(* IEC 61131-3 sources: daoli-st-library/DL_Device (part 23) *)

(* ---- FB_DL_GreaseLubeTimer.st ---- *)
(*
  Name        : FB_DL_GreaseLubeTimer
  Category    : DL_Device
  Version     : 1.0.0
  Purpose     : 加脂保养窗：运行小时数与动作循环数双触发（任一达限即报「该加脂」，先到先报），保养完成后复位清零重计；/ Grease lubrication window: running hours and cycle count both trigger (whichever reaches its limit first reports), cleared and restarted after maintenance
  溯源        : 借 t2-8 ◐/自研 的分类/参数域组织，clean-room 实现
  Boundary    : ① 组态闸：小时限/循环限任一 < 0 → 锁存故障（两限可独立为 0 表示该源不触发，但不可为负）；
                ② 运行小时用 1 s 自复位 TON 节拍累计（IN 串 eRun 相位 + bRunning，R188/族③），段 0 无 IF 包裹；
                ③ 双触发独立判据独立归因（R190）：eHoursFirst / eCyclesFirst 各自成因，同拍同到按小时优先归因（不共用成员）；
                ④ 秒计数饱和累加（R28 防回绕），循环数沿计数净额 +1 饱和；
                ⑤ bLubeDue 锁存至复位沿或 bLubeDone 沿（保养完成脉冲，唯一业务清零路径）；
                ⑥ 本件只报保养到期，不执行加脂动作（属主边界）。
*)
TYPE E_DL_GltState :
(
    eIdle  := 0,                             (* 未使能 / Disabled *)
    eRun   := 10,                            (* 保养窗计时计数运行 / Accumulating *)
    eFault := 90                             (* 故障锁存相 / Fault latched *)
);
END_TYPE

TYPE E_DL_GltCause :
(
    eNone        := 0,                       (* 无故障成因 / No cause *)
    eCfgIllegal  := 1,                       (* 组态非法：时限/循环限越域 / Illegal config *)
    eHoursFirst  := 2,                       (* 运行小时先达限（先到先报） / Hours limit reached first *)
    eCyclesFirst := 3,                       (* 动作循环先达限（先到先报） / Cycles limit reached first *)
    ePhaseBad    := 4                        (* 非法相位兜底 / Illegal phase fallback *)
);
END_TYPE

FUNCTION_BLOCK FB_DL_GreaseLubeTimer
VAR_INPUT
    bRunning   : BOOL := FALSE;              (* 设备运行电平（运行小时累计门控）[-] / Equipment running level *)
    bCyclePulse: BOOL := FALSE;              (* 动作循环脉冲（上升沿计一次）[-] / One action-cycle pulse *)
    fHoursLimit: REAL := 2000.0;             (* 运行小时触发限，域 >= 0（0 = 该源禁用）[h] / Hours trigger limit, >= 0 *)
    nCycleLimit: UDINT := 100000;            (* 循环数触发限，域 >= 0（0 = 该源禁用）[次] / Cycle trigger limit, >= 0 *)
    bLubeDone  : BOOL := FALSE;              (* 保养完成脉冲（业务清零路径，重开保养窗）[-] / Maintenance done pulse *)
    bEnable    : BOOL := TRUE;               (* 使能 [-] / Enable *)
    bReset     : BOOL := FALSE;              (* 复位命令，上升沿清累计与故障 [-] / Reset command *)
END_VAR
VAR_OUTPUT
    fRunHours  : REAL;                       (* 累计运行小时（窗内）[h] / Accumulated running hours *)
    nCycles    : UDINT;                      (* 累计动作循环数（窗内，饱和）[次] / Accumulated cycles, saturated *)
    bLubeDue   : BOOL;                       (* 加脂到期锁存（复位沿或保养完成沿清）[-] / Lubrication due latched *)
    eState     : E_DL_GltState;              (* 状态出口 / State outlet *)
    eCause     : E_DL_GltCause;              (* 成因出口（R190 双触发独立归因） / Cause outlet *)
    bError     : BOOL;                       (* 故障锁存标志 [-] / Fault latch flag *)
END_VAR
VAR
    _eState  : E_DL_GltState := E_DL_GltState.eIdle;     (* 内部相位（CASE 唯一写入目标） / Internal phase *)
    _eCause  : E_DL_GltCause := E_DL_GltCause.eNone;     (* 故障成因锁存量 / Latched cause *)
    rtCycle  : R_TRIG;                       (* 循环脉冲沿实例，段 0 无条件调用 / Cycle pulse edge *)
    rtLube   : R_TRIG;                       (* 保养完成沿实例，段 0 无条件调用 / Lube-done edge instance *)
    rtReset  : R_TRIG;                       (* 复位沿实例，段 0 无条件调用 / Reset edge instance *)
    tonTick  : TON;                          (* 1 s 节拍计时器（自复位，IN 串相位 + 运行电平） / 1 s tick timer *)
    _bFault  : BOOL;                         (* 故障锁存位 / Latched fault bit *)
    _bCfgBad : BOOL;                         (* 组态非法当拍量 / Illegal config this scan *)
    _fSec    : REAL;                         (* 窗内累计运行秒数（节拍累加）[s] / Accumulated seconds *)
    _fHoursI : REAL;                         (* 运行小时中间量（秒→小时换算）[h] / Hours intermediate *)
    _bDueI   : BOOL;                         (* 到期内部量（锁存副本源）[-] / Due internal, source of latch *)
END_VAR
VAR CONSTANT
    DL_GLT_EPS    : REAL  := 1.0E-6;         (* 判零容差 [-] / Epsilon *)
    DL_GLT_CNTMAX : UDINT := 4294967295;     (* 循环计数饱和上限（R28）[-] / Cycle count saturation cap *)
    DL_GLT_SECMAX : REAL  := 3.0E9;          (* 秒累计上限（防 REAL 有效位耗尽，约 95 年）[s] / Seconds accumulation cap *)
    DL_GLT_H2S    : REAL  := 3600.0;         (* 小时→秒换算常量（乘性常量）[-] / Hours to seconds factor *)
END_VAR

(* —— 段 0：当拍判据派生 + 实例无条件刷新（R228A；R_TRIG/TON 全在段 0，无 IF 包裹） —— *)
_bCfgBad := (fHoursLimit < 0.0) OR (nCycleLimit < 0);                          (* 两触发限非负闸（0 = 禁用该源，合法） / Limits non-negative gates *)
rtCycle(CLK := bCyclePulse);                                                   (* 循环沿每拍必调 / Cycle edge every scan *)
rtLube(CLK := bLubeDone);                                                      (* 保养完成沿每拍必调 / Done edge every scan *)
rtReset(CLK := bReset);                                                        (* 复位沿每拍必调 / Reset edge every scan *)
tonTick(IN := (_eState = E_DL_GltState.eRun) AND bRunning AND NOT tonTick.Q, PT := T#1S);   (* 1 s 节拍自复位（R188）+ eRun 相位与运行电平闸 / 1 s tick with phase and run gates *)

(* —— 段 1：单拍量预清零（R107） —— *)
_bDueI := FALSE;                                                               (* 到期内部量预清（判据拍重算） / Due internal preset *)
_fHoursI := 0.0;                                                               (* 小时中间量预清 / Hours intermediate preset *)

(* —— 段 2：复位沿处理（作用域：清故障 + 清累计 + 清到期 + 迁 eIdle，R283 逐项声明） —— *)
IF rtReset.Q THEN
    _bFault := FALSE;                                                          (* 清故障锁存 / Clear fault *)
    _eCause := E_DL_GltCause.eNone;                                            (* 清成因 / Clear cause *)
    _fSec := 0.0;                                                              (* 清秒累计 / Clear seconds *)
    nCycles := 0;                                                              (* 清循环计数出口 / Clear cycles outlet *)
    bLubeDue := FALSE;                                                         (* 清到期锁存出口 / Clear due outlet *)
    _eState := E_DL_GltState.eIdle;                                            (* 迁未使能相 / Back to idle *)
END_IF

(* —— 段 3：组态故障锁存（锁存至复位沿，R189） —— *)
IF _bCfgBad AND NOT _bFault THEN
    _bFault := TRUE;                                                           (* 锁存故障位 / Latch fault *)
    _eCause := E_DL_GltCause.eCfgIllegal;                                      (* 成因：组态非法 / Cause: illegal config *)
    _eState := E_DL_GltState.eFault;                                           (* 同步迁故障相 / Migrate to fault *)
END_IF

(* —— 段 4：CASE 主状态机（ELSE 兜底迁 eFault，红线 6） —— *)
CASE _eState OF
    E_DL_GltState.eIdle:                                                       (* 未使能：不累计，出口确定值 / Disabled *)
        _fSec := 0.0;                                                          (* 失能清秒累计（防隐性回夹） / Clear seconds *)
        fRunHours := 0.0;                                                      (* 失能清小时出口 / Clear hours outlet *)
        nCycles := 0;                                                          (* 失能清循环出口 / Clear cycles outlet *)
        bLubeDue := FALSE;                                                     (* 失能清到期出口 / Clear due outlet *)
        IF bEnable AND NOT _bFault THEN
            _eState := E_DL_GltState.eRun;                                     (* 使能进入累计 / Enter accumulating *)
        END_IF
    E_DL_GltState.eRun:                                                        (* 累计相：小时 + 循环双源 / Accumulating *)
        IF NOT bEnable THEN
            _eState := E_DL_GltState.eIdle;                                    (* 失能回未使能 / Back to idle *)
        ELSE
            IF rtLube.Q THEN                                                   (* 保养完成沿：业务清零重开窗（唯一业务清零路径） / Done edge: clear and reopen window *)
                _fSec := 0.0;                                                  (* 清秒累计 / Clear seconds *)
                nCycles := 0;                                                  (* 清循环计数 / Clear cycles *)
                bLubeDue := FALSE;                                             (* 清到期锁存 / Clear due latch *)
                _eCause := E_DL_GltCause.eNone;                                (* 成因复位 / Cause reset *)
            END_IF
            IF tonTick.Q THEN                                                  (* 1 s 节拍到点：秒累计 +1 / Tick elapsed: +1 second *)
                IF _fSec < DL_GLT_SECMAX THEN
                    _fSec := _fSec + 1.0;                                      (* 秒累计（饱和防有效位耗尽，R28） / Seconds accumulate, capped *)
                END_IF
            END_IF
            IF rtCycle.Q THEN                                                  (* 动作循环沿：循环计数 +1 / Cycle edge: +1 *)
                IF nCycles < DL_GLT_CNTMAX THEN
                    nCycles := nCycles + 1;                                    (* 循环计数净额 +1（饱和防回绕） / Net +1, saturated *)
                END_IF
            END_IF
            _fHoursI := _fSec / DL_GLT_H2S;                                    (* 秒→小时换算（除子为常量）[h] / Seconds to hours *)
            fRunHours := _fHoursI;                                             (* 小时出口 / Hours outlet *)
            IF (fHoursLimit > DL_GLT_EPS) AND (_fHoursI >= fHoursLimit) THEN   (* 小时源触发（源限 0 = 禁用不判） / Hours trigger *)
                _bDueI := TRUE;                                                (* 到期内部量置位 / Due set *)
                IF NOT bLubeDue THEN
                    _eCause := E_DL_GltCause.eHoursFirst;                      (* 先到先报：小时源归因（R190） / Hours-first attribution *)
                END_IF
            END_IF
            IF (nCycleLimit > 0) AND (nCycles >= nCycleLimit) THEN             (* 循环源触发（源限 0 = 禁用不判） / Cycle trigger *)
                _bDueI := TRUE;                                                (* 到期内部量置位 / Due set *)
                IF NOT bLubeDue THEN
                    _eCause := E_DL_GltCause.eCyclesFirst;                     (* 先到先报：循环源归因（小时已报则保持小时归因） / Cycles-first attribution *)
                END_IF
            END_IF
            IF _bDueI THEN
                bLubeDue := TRUE;                                              (* 到期锁存（复位沿/保养沿清） / Latch due *)
            END_IF
        END_IF
    E_DL_GltState.eFault:                                                      (* 故障相：冻结保持末值，仅复位沿出 / Fault *)
        ;                                                                      (* 锁存回放（R28） / Replay from latch *)
    ELSE                                                                       (* 非法相位兜底迁安全态 / Illegal phase fallback *)
        _eState := E_DL_GltState.eFault;                                       (* 迁故障相 / To fault *)
        _bFault := TRUE;                                                       (* 同步锁存 / Latch *)
        _eCause := E_DL_GltCause.ePhaseBad;                                    (* 成因：非法相位 / Cause: illegal phase *)
END_CASE

(* —— 段 5：出口映射（bError/eState 同源，R191） —— *)
bError := _bFault;                                                             (* 故障标志镜像 / Fault flag mirror *)
eState := _eState;                                                             (* 状态出口 / State outlet *)
eCause := _eCause;                                                             (* 成因出口 / Cause outlet *)
END_FUNCTION_BLOCK

(* ---- FB_DL_HealthAggregator.st ---- *)
//==============================================================================
// 功能块：FB_DL_HealthAggregator ｜ 中文名称：多源 NE107 健康聚合仲裁
// 所属子库：DL_Device ｜ 版本：v1.0.0 ｜ 兼容：CODESYS V3.5+ / TwinCAT 3 / 汇川 InoProShop
// 功能描述：多源 NE107 健康态聚合仲裁件——对至多 16 路健康源按枚举序号
//           "最差者胜"（编号最小者优先）聚合出总健康态，并给出最差源
//           下标与失效/维护两级计数。HMI 顶部健康横幅的单一事实源。
// 开源溯源 (Origin)：道莅 clean-room 防御性实现
// 单位表：健康态[—]（E_DL_Ne107Status 序号）／源路数[路]／下标[路]
// 错误码表：16#0003_017A 信息级（源数 > 16 已钳位 16 照常仲裁，不置
//           bError）/ 16#0003_017B 信息级（全部源均为 eUnknown，输出
//           eUnknown 是合法结论非错误）/ 16#0003_0348 故障级（源数为 0，
//           无可仲裁对象，置 bError）/ 16#0003_0349 预留禁用（不得挪用）/
//           16#0003_034A 故障级兜底（置 bError，本件纯当拍仲裁无状态机，
//           兜底码保留给未来状态化扩展误用拦截）
// 状态机：N/A（纯当拍仲裁，无状态机、无迟滞、无跨拍锁存；聚合无迟滞，
//           调用方如需防抖自行组合 FB_DL_SignalDebounce 后再接入 aHealth）
// 边界行为：① uSourceCount > 16 → 钳 16 + 信息 017A，数组访问一律有
//           uIdx <= 16 二次闸（字面量上界与 DL_HEALTH_MAX 一致性由本件
//           承担验证责任，两处同源 16）；② uSourceCount = 0 → 故障 0348、
//           eOverall := eUnknown、bValid := FALSE；③ 全部源 eUnknown →
//           输出 eUnknown + 信息 017B（合法结论，不置故障）；④ bArbitrate
//           = FALSE → 本拍不仲裁，eOverall := eUnknown、bValid := FALSE
//           （不冻结旧值，横幅显示"未仲裁"口径）；⑤ 数组访问下标越界
//           理论不可能（钳位 + 二次闸双保险），仍以防御闸兜底。
// 依赖纪律：仅 Standard.library + 同库契约 E_DL_Ne107Status（属主
//           I_DL_DeviceHealth.st，只引用不重声明，R70）；零同层调用。
// 修订历史：v1.0.0 2026-11-17 首版（R23 派单 · T2-8 NE107 待挖项落地）
//==============================================================================

(*------------------------------------------------------------------------------
 * 调用示例：HMI_Health(IN := aHealth, uSourceCount := uN, bArbitrate := TRUE);
 *   HMI 横幅：IF fbHMI.eOverall <= E_DL_Ne107Status.eCheckFunction THEN
 *                 红色横幅; ELSIF fbHMI.eOverall <= eOutOfSpec THEN 黄色; 其余态类似降档
 *   仅当 bValid = TRUE 且 eErr 属信息级（017A/017B）时聚合结果可用于
 *   画面/报表；eErr = 0348 时横幅显示"组态错误"。
 *-----------------------------------------------------------------------------*)
FUNCTION_BLOCK FB_DL_HealthAggregator
VAR_INPUT
    aHealth     : ARRAY[1..16] OF E_DL_Ne107Status; // 各源健康态 [—]，下标 1..16，超编路填 eUnknown / Health status per source, index 1..16, over-count lanes fill eUnknown
    uSourceCount: UINT;                     // 实际源数 [路]，有效域 0..16，> 16 钳位照仲裁 / Actual source count [lanes], 0..16, clamped above
    bArbitrate  : BOOL;                     // 仲裁使能 [—]，FALSE = 本拍不仲裁输出 eUnknown / Arbitration enable, FALSE = skip and report eUnknown
END_VAR
VAR_OUTPUT
    eOverall    : E_DL_Ne107Status;         // 聚合结果 [—]，编号最小者优先即最差者胜 / Aggregated status, lowest ordinal wins, the worst prevails
    uWorstIdx   : UINT;                     // 最差源下标 [路]，0 = 无（未仲裁或源数为 0） / Worst source index [lanes], 0 = none
    uFailCount  : UINT;                     // eFailure 源计数 [路] / Count of eFailure sources [lanes]
    uMaintCount : UINT;                     // eMaintenanceReq 源计数 [路] / Count of eMaintenanceReq sources [lanes]
    eErr        : UDINT;                    // 错误码，0 = 无错 / Error code, 0 = no error
    bError      : BOOL;                     // 故障级标志，仅故障级错误置位 / Fault-class flag, set only on fault-level codes
    bValid      : BOOL;                     // 输出可用标志 / Outputs usable flag
END_VAR
VAR CONSTANT
    DL_HEALTH_MAX : UINT := 16;             // 数组上界 [路]，与接口字面量上界 16 同源，改动须同步 / Array ceiling [lanes], same source as the literal bound 16, change both together
END_VAR
VAR
    uCountEff   : UINT;                     // 钳位后的生效源数 [路] / Effective clamped source count [lanes]
    uIdx        : UINT;                     // 扫描循环下标 [路] / Scan loop index [lanes]
    eWorst      : E_DL_Ne107Status;         // 当前最差态暂存 [—] / Staged worst status so far
    uWorstStaged: UINT;                     // 当前最差源下标暂存 [路] / Staged worst index so far
END_VAR

(*------------------------------------------------------------------------------
 * 段 1｜每拍预置：纯当拍仲裁，全部输出每拍重算，无保持量、无首扫分支
 *      Pure per-scan arbitration, every output recomputed, no held state
 *-----------------------------------------------------------------------------*)
eOverall     := E_DL_Ne107Status.eUnknown;   // 聚合结果预置未知 / Aggregated result preset unknown
uWorstIdx    := 0;                           // 最差源下标预置无 / Worst index preset to none
uFailCount   := 0;                           // 失效计数清零 / Failure count cleared
uMaintCount  := 0;                           // 维护计数清零 / Maintenance count cleared
eErr         := 16#0000_0000;                // 错误码每拍重算 / Error code recomputed
bError       := FALSE;                       // 故障标志每拍重算 / Fault flag recomputed
bValid       := FALSE;                       // 可用标志每拍重算 / Usable flag recomputed
uCountEff    := 0;                           // 生效源数预置零 / Effective count preset zero
eWorst       := E_DL_Ne107Status.eUnknown;   // 最差态暂存预置未知 / Staged worst preset unknown
uWorstStaged := 0;                           // 最差下标暂存预置零 / Staged worst index preset zero

(*------------------------------------------------------------------------------
 * 段 2｜仲裁使能与源数闸门（0 → 故障；> 16 → 钳位 + 信息）
 *      Arbitration enable and source-count gates
 *-----------------------------------------------------------------------------*)
IF NOT bArbitrate THEN
    eOverall := E_DL_Ne107Status.eUnknown;  // 未仲裁口径：输出未知 / Not arbitrating, report unknown
    RETURN;                                 // bValid 保持 FALSE / bValid stays FALSE
END_IF
IF uSourceCount = 0 THEN
    eOverall := E_DL_Ne107Status.eUnknown;  // 无可仲裁对象 / Nothing to arbitrate
    eErr   := 16#0003_0348;                 // 故障级：源数为 0 / Fault: zero sources
    bError := TRUE;                         // 置故障标志（R45 配对） / Raise the fault flag
    bValid := FALSE;                        // 输出不可用 / Outputs unusable
    RETURN;
END_IF
IF uSourceCount > DL_HEALTH_MAX THEN
    uCountEff := DL_HEALTH_MAX;             // 源数钳位到 16 路照仲裁 / Count clamped to 16 lanes
    eErr := 16#0003_017A;                   // 信息级：源数已钳位（不置 bError） / Info: count clamped, no fault flag
ELSE
    uCountEff := uSourceCount;              // 合法源数原值生效 / Valid count applied as-is
END_IF

(*------------------------------------------------------------------------------
 * 段 3｜最差者胜扫描：编号最小者优先（eFailure=0 最差，eOk=40 最好）；
 *       下标访问带 uIdx <= 16 二次闸（R 二次闸纪律），并统计两级计数
 *       Worst-prevails scan with the secondary index gate and two counters
 *-----------------------------------------------------------------------------*)
FOR uIdx := 1 TO uCountEff DO
    IF uIdx <= DL_HEALTH_MAX THEN           // 二次闸：越界访问结构性不可能 / Secondary gate, out-of-bounds structurally impossible
        IF aHealth[uIdx] < eWorst THEN      // 序号更小 = 更差 / Lower ordinal means worse
            eWorst := aHealth[uIdx];        // 更新最差态 / Update the worst status
            uWorstStaged := uIdx;           // 记录最差源下标 / Record the worst source index
        END_IF
        IF aHealth[uIdx] = E_DL_Ne107Status.eFailure THEN
            uFailCount := uFailCount + 1;   // 失效源计数递增 / Failure counter increment
        END_IF
        IF aHealth[uIdx] = E_DL_Ne107Status.eMaintenanceReq THEN
            uMaintCount := uMaintCount + 1; // 维护源计数递增 / Maintenance counter increment
        END_IF
    END_IF
END_FOR

(*------------------------------------------------------------------------------
 * 段 4｜出口：全未知声明 + 可用性
 *      Outlet: all-unknown notice and usability
 *-----------------------------------------------------------------------------*)
eOverall  := eWorst;                        // 聚合结果出口 / Aggregated result outlet
uWorstIdx := uWorstStaged;                  // 最差源下标出口 / Worst index outlet
IF eWorst = E_DL_Ne107Status.eUnknown THEN
    eErr := 16#0003_017B;                   // 信息级：全部源未知，合法结论（不置 bError） / Info: all sources unknown, a legal conclusion
END_IF
bValid := TRUE;                             // 输出可用（含信息级情形） / Outputs usable, including info-level cases
END_FUNCTION_BLOCK

(* ---- FB_DL_HealthStatusArbiter.st ---- *)
(*
  Name        : FB_DL_HealthStatusArbiter
  Category    : DL_Device
  Version     : 1.0.0
  Purpose     : 多源 NE107 健康仲裁聚合：N 路健康枚举逐件直比最差胜出（仅已知源参与），聚合出口单一健康态；/ Multi-source NE107 health arbitration: N health status entries compared item-wise with the worst known winning, aggregated into a single health outlet
  溯源        : 借 t2-8 NE107/ISA-18.2 的分类/参数域组织，clean-room 实现
  依赖声明    : 引用 E_DL_Ne107Status（唯一属主 DL_Device 契约件 I_DL_DeviceHealth），不重造枚举；
                该枚举数值即优先级：数值最小最差（eFailure = 0 最差，eOk = 40，eUnknown = 99 不参与仲裁）。
  Boundary    : ① 源计数越界钳 NMAX（8），负数/零计数聚合出 eUnknown 且来源序号出口 0；
                ② 最差态判定为数值直比取最小（编号即优先级），逐件遍历无排序无锁存；
                ③ 单路 eUnknown 不抬高也不拉低聚合结论（仅已知源参与），全部未知时聚合出 eUnknown；
                ④ 仲裁为纯组合重算（无状态机、无锁存），每拍全量重判防陈旧（本件按边界④不设相位机）；
                ⑤ 出口与 I_DL_DeviceHealth 六态契约同源（E_DL_Ne107Status），不重造枚举；
                ⑥ 零外部全局、零物理地址，纯函数式聚合可跨平台移植。
*)
FUNCTION_BLOCK FB_DL_HealthStatusArbiter
VAR_INPUT
    aHealth : ARRAY[1..8] OF E_DL_Ne107Status;   (* 各源 NE107 健康态（六态契约同源）[-] / Health status per source *)
    nCount  : INT := 8;                      (* 参与仲裁源计数，域 1..8 [路] / Source count in arbitration *)
END_VAR
VAR_OUTPUT
    eAgg    : E_DL_Ne107Status;              (* 聚合健康态出口（最差胜出）[-] / Aggregated health outlet *)
    nWorstSrc: INT;                          (* 最差来源序号（1 基，0 = 无已知源）[-] / Worst source index *)
    nKnown  : INT;                           (* 已知源计数（诊断）[路] / Known source count *)
END_VAR
VAR CONSTANT
    DL_HSA_NMAX   : INT := 8;                (* 源数容量上限（钳位）[路] / Source capacity limit *)
END_VAR
VAR
    _eWorst : E_DL_Ne107Status := E_DL_Ne107Status.eUnknown;   (* 当前最差态（哨兵 = 未知，枚举直存不转整数） / Current worst status *)
    _nKnown : INT;                           (* 已知源计数累加量 [路] / Known source accumulator *)
    _i      : INT;                           (* 生效源计数（钳位后）[路] / Effective source count *)
    _j      : INT;                           (* 遍历游标 [路] / Loop cursor *)
END_VAR

(* —— 段 1：出口预清（组合确定性出口，无陈旧，R107） —— *)
eAgg := E_DL_Ne107Status.eUnknown;                       (* 聚合出口预置未知 / Agg outlet preset unknown *)
nWorstSrc := 0;                                          (* 最差来源序号预置 0 / Worst source preset zero *)
_nKnown := 0;                                            (* 已知源计数清零 / Known count clear *)
_eWorst := E_DL_Ne107Status.eUnknown;                    (* 最差态预置哨兵（未遇到已知源） / Worst preset sentinel *)
nKnown := 0;                                             (* 已知源计数出口预清 / Known count outlet preset *)

(* —— 段 2：源计数域闸 + 钳位（边界①） —— *)
IF (nCount < 1) OR (nCount > DL_HSA_NMAX) THEN
    _i := DL_HSA_NMAX;                                   (* 越界钳上限（含负数与零保护） / Clamp to capacity *)
ELSE
    _i := nCount;                                        (* 域内直用 / In domain direct *)
END_IF

(* —— 段 3：逐件直比仲裁（枚举有序比较，最小 = 最差胜出，边界②③；FOR 有界无死循环） —— *)
FOR _j := 1 TO _i DO
    IF aHealth[_j] <> E_DL_Ne107Status.eUnknown THEN     (* 未知源不参与仲裁（边界③） / Unknown source skipped *)
        _nKnown := _nKnown + 1;                          (* 已知源计数累加 / Known count accumulate *)
        IF aHealth[_j] < _eWorst THEN                    (* 枚举有序直比取最小 = 最差（编号即优先级） / Enum ordered compare, min wins *)
            _eWorst := aHealth[_j];                      (* 更新最差态 / Update worst *)
            nWorstSrc := _j;                             (* 记录最差来源序号 / Record worst source *)
        END_IF
    END_IF
END_FOR
nKnown := _nKnown;                                       (* 已知源计数出口 / Known count outlet *)

(* —— 段 4：聚合出口映射（全未知 → eUnknown 哨兵保持，边界③④） —— *)
IF _eWorst <> E_DL_Ne107Status.eUnknown THEN
    eAgg := _eWorst;                                     (* 最差态回映射聚合出口 / Worst to aggregate outlet *)
END_IF
END_FUNCTION_BLOCK

(* ---- FB_DL_HeaterBankLoadBalance.st ---- *)
(*
    FB_DL_HeaterBankLoadBalance —— 加热器组负载均衡选主
    ------------------------------------------------------------------
    分类      : DL_Device / Thermal
    前缀      : FB_DL_
    版本      : 1.0.0
    溯源      : clean-room 自有实现；仅借鉴「按累计工时轮换主用」的公开运维常识语义，
                未复制任何闭源厂商源码，码位 100% 自有
    平台      : 纯 IEC 61131-3，CODESYS V3.5+ / TwinCAT 3 / InoProShop / Machine Expert 通用
    作者      : 道莅代码库 · PLC编程专家（R76 冲刺批 C3 · #2）
    ------------------------------------------------------------------
    功能说明  : N 路加热器（rN 钳位 2..8）按累计运行工时选主：每拍从可用通道
                （健康 AND 投运允许 AND 工时有限）中选累计工时最小者为主通道，
                工时相同（容差内）按通道号小者优先；主通道故障自动顺延次小工时通道；
                超温（fTemp > fDerateTh）整组降额占空比至 fDerateDuty，带滞回恢复。
                边界：只产出主通道号与各通道占空比指令，不直接驱动 DO/PWM 硬件，
                工时累计由上位系统维护、本件只读。
    R6 口径    : 主状态机 E_DL_HeatBalState（eIdle/eRun/eFault）为 ENUM+CASE+ELSE，
                ELSE 置 16#0005_1E06 并回 eFault；选主逻辑为无跨拍状态驻留的判据链
                （FOR 升序遍历 + 严格小于 + 容差，天然满足「同工时通道号小者优先」），
                判据链等价 CASE 的兜底由「全通道不可用 → 1E01」分支承担。
    错误码    : 16#0005_1E00 参数非法（占空比出 [0,1] / 滞回为负 / 降额阈不大于滞回）——故障级
                16#0005_1E01 全部通道不可用，无主可选——故障级，锁存至复位沿
                16#0005_1E02 主通道故障顺延次小工时通道——信息级，顺延拍单发
                16#0005_1E03 超温降额激活——信息级，降额期间持续发布
                16#0005_1E04 通道工时非有限，按不可用剔除该通道——信息级，条件存在即发布
                16#0005_1E05 温度采样非有限，保持降额占空比（安全侧）——故障级，条件级不锁存
                16#0005_1E06 CASE 落 ELSE 兜底——故障级
    码位总账  : 16#0005_1E00..1E06 全部定义并使用，无空悬码位；
                信息级码同拍多发时以后赋值者可见（1E05 优先级最高，最后赋值）
    状态机    : eIdle --bBankEnable 且参数合法--> eRun；eRun 内全通道不可用 → eFault
                （1E01 锁存，bReset 上升沿复位）；1E05 为条件级故障不转 eFault、
                保持降额占空比继续选主；1E00 门禁非法直接转 eFault。
    防御口径  : 工时比较用绝对容差 DL_HB_EPS（工时差归一无需除法，本件无除法运算，
                分母不存在）；通道下标一律 1..8 硬界内，nMaster 只能取自
                1..nEff（nEff 已钳位 2..8），占空比映射用等值比较杜绝越界；
                非有限判定按 NaN f<>f、±Inf (f-f)<>(f-f)。
    修订记录  : 2026-11-23 v1.0.0 首次入库（R76 冲刺批 C3 · #2）
*)
TYPE E_DL_HeatBalState :
(
    eIdle  := 0,   // 待机，整组未投运，占空比全零 / idle, bank off, all duties zero
    eRun   := 10,  // 运行，每拍重算选主与占空比 / running, master selection and duties recomputed every scan
    eFault := 20   // 故障，主通道清零、占空比全零，锁存码等复位 / fault, master cleared, duties zero, code latched for reset
);
END_TYPE

FUNCTION_BLOCK FB_DL_HeaterBankLoadBalance
VAR_INPUT
    rN          : INT;                     // 配置通道数，钳位到 2..8 / configured channel count, clamped to 2..8
    aHours      : ARRAY[1..8] OF LREAL;    // 各通道累计运行工时 [h]，上位维护、本件只读 / accumulated run hours [h] per channel, maintained upstream, read-only here
    aHealthy    : ARRAY[1..8] OF BOOL;     // 各通道健康标志，TRUE = 可用 / per-channel health flag, TRUE = available
    aEnabled    : ARRAY[1..8] OF BOOL;     // 各通道投运允许，TRUE = 参与选主 / per-channel enable, TRUE = joins the selection
    fTemp       : REAL;                    // 加热组温度采样 [°C] / bank temperature sample [°C]
    fDerateTh   : REAL := 80.0;            // 超温降额阈值 [°C]，必须大于滞回 / derate threshold [°C], must exceed the hysteresis
    fDerateHys  : REAL := 2.0;             // 降额恢复滞回 [°C]，非负 / derate release hysteresis [°C], non-negative
    fDerateDuty : REAL := 0.5;             // 降额占空比 [0..1] / derated duty cycle [0..1]
    fNomDuty    : REAL := 1.0;             // 正常占空比 [0..1] / nominal duty cycle [0..1]
    bBankEnable : BOOL;                    // 整组投运命令 / bank enable command
    bReset      : BOOL;                    // 故障复位请求，上升沿生效 / fault reset request, edge-active
END_VAR
VAR_OUTPUT
    nMaster     : INT;                     // 当前主通道号 1..8，0 = 无主 / current master channel 1..8, 0 = none
    aDuty       : ARRAY[1..8] OF REAL;     // 各通道占空比指令 [0..1]，非主通道恒 0 / duty command [0..1] per channel, non-master channels are 0
    bDerated    : BOOL;                    // 整组降额标志 / bank derated flag
    eState      : E_DL_HeatBalState;       // 当前状态镜像输出 / current state mirror output
    nErrCode    : UDINT;                   // 错误码，0 = 无错；信息级随条件发布、故障级锁存回放 / error code, 0 = none; info codes conditional, fault codes latched
    bError      : BOOL;                    // 故障级标志，仅故障级码置位 / fault-class flag, raised only by fault-class codes
    bValid      : BOOL;                    // 输出可用标志，= NOT bError / outputs valid flag, equals NOT bError
END_VAR
VAR
    _eState      : E_DL_HeatBalState;      // 当前状态 / current state
    _uErrLatch   : UDINT;                  // 故障码锁存副本，故障态每拍回放 / latched fault code republished inside the fault state
    rtReset      : R_TRIG;                 // 复位上升沿检测 / reset rising-edge detector
    _nEff        : INT;                    // 钳位后的有效通道数 2..8 / effective channel count clamped to 2..8
    _nBest       : INT;                    // 本拍选出的主通道号 / master channel selected this scan
    _nMasterPrev : INT;                    // 上一拍主通道号，顺延观测用 / previous-scan master channel for the fallback observation
    _fBest       : LREAL;                  // 本拍最小工时 [h] / smallest hours found this scan [h]
    _fDuty       : REAL;                   // 本拍主通道占空比 [0..1] / master duty this scan [0..1]
    _i           : INT;                    // FOR 循环变量，1..8 硬界 / FOR loop index within the hard 1..8 bounds
    _bAvail      : BOOL;                   // 通道可用临时量 / per-channel availability scratch
    _bParOk      : BOOL;                   // 参数门禁结果 / parameter gate result
    _bTempBad    : BOOL;                   // 温度采样非有限标志 / non-finite temperature flag
    _bDerateLatch : BOOL;                  // 降额滞回锁存 / derate hysteresis latch
END_VAR
VAR CONSTANT
    DL_HB_EPS   : LREAL := 1.0E-9;         // 工时比较容差 [h]，容差内视为同工时 / hours comparison tolerance [h], inside it hours count as equal
    DL_HB_TOL   : REAL  := 1.0E-6;         // 占空比域比较容差 [无量纲] / duty domain comparison tolerance [dimensionless]
    DL_HB_ZERO  : REAL  := 0.0;            // 零占空比 [0..1] / zero duty [0..1]
    DL_HB_ONE   : REAL  := 1.0;            // 满占空比域上界 [0..1] / full-duty domain upper bound [0..1]
    DL_HB_CHMIN : INT   := 2;              // 通道数下限 / channel count lower bound
    DL_HB_CHMAX : INT   := 8;              // 通道数上限（数组硬界）/ channel count upper bound, the array hard bound
END_VAR

// 段 1｜边缘检测无条件周期刷新（R7：严禁放入 IF / CASE；本件无 TON）
// segment 1, edge detector refreshed unconditionally, never inside IF/CASE; no TON in this FB
rtReset(CLK := bReset);

// 段 2｜输出与错误状态预置；故障态从锁存副本回放（R45 配对）
// segment 2, preset outputs and error status; the fault state replays from the latch
nMaster := 0;                              // 预置无主 / preset no master
bDerated := FALSE;                         // 预置未降额 / preset not derated
nErrCode := 0;                             // 预置无错误码 / preset no error code
bError := FALSE;                           // 预置无故障标志 / preset no fault flag
bValid := TRUE;                            // 预置输出可用 / preset outputs valid
IF _eState = E_DL_HeatBalState.eFault THEN
    nErrCode := _uErrLatch;                // 重发布锁存故障码 / republish the latched fault code
    bError := TRUE;                        // 故障态恒置故障标志 / fault flag stays raised in the fault state
    bValid := FALSE;                       // 故障态输出不可信 / outputs not valid in the fault state
END_IF

// 段 3｜参数门禁与通道数钳位：rN 钳位属正常行为不报错，其余非法即锁存 1E00 转 eFault
// segment 3, parameter gate and channel clamp; rN clamping is normal behaviour, other violations latch 1E00 and jump to eFault
_nEff := rN;                               // 取配置通道数 / take the configured channel count
IF _nEff < DL_HB_CHMIN THEN
    _nEff := DL_HB_CHMIN;                  // 钳到下限 2 / clamp to the lower bound 2
END_IF
IF _nEff > DL_HB_CHMAX THEN
    _nEff := DL_HB_CHMAX;                  // 钳到上限 8（数组硬界）/ clamp to the upper bound 8, the array hard bound
END_IF
_bParOk := (fDerateDuty > (DL_HB_ZERO - DL_HB_TOL)) AND (fDerateDuty < (DL_HB_ONE + DL_HB_TOL))
       AND (fNomDuty > (DL_HB_ZERO - DL_HB_TOL)) AND (fNomDuty < (DL_HB_ONE + DL_HB_TOL))
       AND (fDerateHys > (DL_HB_ZERO - DL_HB_TOL)) AND (fDerateTh > fDerateHys);
_bTempBad := (fTemp <> fTemp) OR ((fTemp - fTemp) <> (fTemp - fTemp)); // 温度 NaN/±Inf 判定 / temperature NaN or infinite
IF (NOT _bParOk) AND (_eState <> E_DL_HeatBalState.eFault) THEN
    _uErrLatch := 16#0005_1E00;            // 锁存参数非法码 / latch the illegal parameter code
    nErrCode := 16#0005_1E00;              // 故障级码赋值 3 行内置 bError / fault-class assignment with bError inline
    bError := TRUE;
    bValid := FALSE;
    _eState := E_DL_HeatBalState.eFault;   // 参数不可信直接转故障 / untrusted parameters jump to fault
END_IF

// 段 4｜主状态机：CASE + ELSE 兜底（R6）；选主判据链在 eRun 相内每拍全量重算
// segment 4, main state machine, CASE with ELSE fallback; the selection chain inside eRun is recomputed fully every scan
CASE _eState OF
E_DL_HeatBalState.eIdle:
    // 拍 N 进入：复位或未投运；本拍行为：占空比全零（预置已清）；拍 N+1 转出：投运且参数合法 → eRun
    // entered after reset or when off; duties stay zero via the preset; exits to eRun on bank enable with legal parameters
    IF bBankEnable AND _bParOk THEN
        _bDerateLatch := FALSE;            // 新投运清降额锁存 / clear the derate latch on a fresh start
        _nMasterPrev := 0;                 // 清上一拍主通道观测 / clear the previous-master observation
        _eState := E_DL_HeatBalState.eRun; // 进运行相 / enter the run phase
    END_IF

E_DL_HeatBalState.eRun:
    // 拍 N 进入：投运且参数合法；本拍行为：选主 → 顺延观测 → 超温降额 → 占空比映射；
    // 拍 N+1 转出：全通道不可用 → eFault（1E01）；温度非有限保持本相降额运行（1E05 条件级）
    // entered on enable with legal parameters; per scan: select master, observe fallback, derate, map duties;
    // exits to eFault only when no channel is available (1E01); a non-finite temperature keeps this phase derated (1E05)
    _nBest := 0;                           // 清本拍选主结果 / clear this scan's selection
    _fBest := 0.0;                         // 清最小工时 / clear the smallest hours
    FOR _i := 1 TO _nEff DO
        _bAvail := aHealthy[_i] AND aEnabled[_i]; // 可用 = 健康且投运允许 / available = healthy and enabled
        IF (aHours[_i] <> aHours[_i]) OR ((aHours[_i] - aHours[_i]) <> (aHours[_i] - aHours[_i])) THEN
            _bAvail := FALSE;              // 工时非有限剔除该通道 / exclude the channel on non-finite hours
            nErrCode := 16#0005_1E04;      // 信息级：条件存在即发布，不置 bError / info class, no fault flag
        END_IF
        IF _bAvail THEN
            IF (_nBest = 0) OR (aHours[_i] < (_fBest - DL_HB_EPS)) THEN
                _nBest := _i;              // 严格小于才替换：升序遍历 + 容差保证同工时小号优先 / strict less with tolerance keeps the lower index on ties
                _fBest := aHours[_i];      // 记录当前最小工时 / record the current minimum hours
            END_IF
        END_IF
    END_FOR
    IF (_nMasterPrev >= 1) AND (_nMasterPrev <= _nEff)
       AND ((NOT aHealthy[_nMasterPrev]) OR (NOT aEnabled[_nMasterPrev])) AND (_nBest > 0) THEN
        nErrCode := 16#0005_1E02;          // 信息级：主通道故障已顺延（下标受 _nMasterPrev<=_nEff<=8 保护）/ info: master fell over, index guarded
    END_IF
    IF _nBest = 0 THEN
        _uErrLatch := 16#0005_1E01;        // 锁存全通道不可用码 / latch the no-channel-available code
        nErrCode := 16#0005_1E01;          // 故障级码赋值 3 行内置 bError / fault-class assignment with bError inline
        bError := TRUE;
        bValid := FALSE;
        _nMasterPrev := 0;                 // 清观测防复位后误报顺延 / clear the observation to avoid a false fallback after reset
        _eState := E_DL_HeatBalState.eFault; // 转故障，占空比由预置全零 / go to fault, duties stay zero via the preset
    ELSE
        nMaster := _nBest;                 // 发布主通道号 / publish the master channel
        IF fTemp > fDerateTh THEN
            _bDerateLatch := TRUE;         // 超温进入降额 / enter derate on overtemperature
        ELSIF fTemp < (fDerateTh - fDerateHys) THEN
            _bDerateLatch := FALSE;        // 低于恢复阈退出降额（滞回）/ leave derate under the release threshold
        END_IF
        IF _bDerateLatch THEN
            _fDuty := fDerateDuty;         // 降额占空比 / derated duty
            nErrCode := 16#0005_1E03;      // 信息级：降额期间持续发布 / info class, published while derated
        ELSE
            _fDuty := fNomDuty;            // 正常占空比 / nominal duty
        END_IF
        IF _bTempBad THEN
            nErrCode := 16#0005_1E05;      // 温度非有限码最后赋值，显示优先级最高 / assigned last so it wins the display
            _fDuty := fDerateDuty;         // 安全侧：强制降额占空比 / safe side, force the derated duty
            bError := TRUE;                // 故障级码赋值 3 行内置 bError（条件级不锁存，条件消失自动恢复）/ fault-class trio, conditional not latched
            bValid := FALSE;
            bDerated := TRUE;              // 温度不可信视同降额 / untrusted temperature counts as derated
        END_IF
        FOR _i := 1 TO DL_HB_CHMAX DO
            IF _i = nMaster THEN
                aDuty[_i] := _fDuty;       // 主通道承载占空比（nMaster<=_nEff<=8，等值比较无越界）/ master carries the duty, equality test cannot overrun
            ELSE
                aDuty[_i] := DL_HB_ZERO;   // 非主通道恒零 / non-master channels stay zero
            END_IF
        END_FOR
        bDerated := _bDerateLatch OR bDerated; // 汇总降额标志 / merge the derate flag
        _nMasterPrev := nMaster;           // 更新上一拍主通道观测 / update the previous-master observation
    END_IF

E_DL_HeatBalState.eFault:
    // 拍 N 进入：全通道不可用或参数非法；本拍行为：主通道清零（预置）、占空比全零、锁存码回放；
    // 拍 N+1 转出：bReset 上升沿且参数已合法 → eIdle
    // entered on no-channel or illegal parameters; master cleared via the preset, duties zero, latch replays;
    // exits to eIdle on a reset edge with legal parameters
    IF rtReset.Q AND _bParOk THEN
        _uErrLatch := 0;                   // 清锁存码 / clear the latched code
        _eState := E_DL_HeatBalState.eIdle; // 回待机等投运 / back to idle awaiting enable
    END_IF

ELSE
    // 非法状态拦截：任何未定义枚举值一律锁存兜底码并转故障（R6）
    // illegal-state interception, any undefined enum value latches the fallback code and goes to fault
    _uErrLatch := 16#0005_1E06;            // 锁存兜底码 / latch the fallback code
    nErrCode := 16#0005_1E06;              // 故障级码赋值 3 行内置 bError / fault-class assignment with bError inline
    bError := TRUE;
    bValid := FALSE;
    _eState := E_DL_HeatBalState.eFault;
END_CASE

// 段 5｜状态镜像输出
// segment 5, state mirror output
eState := _eState;                         // 状态镜像输出 / state mirror output

END_FUNCTION_BLOCK

(* ---- FB_DL_HeaterBreakDetect.st ---- *)
(*==============================================================================
 * 组件名称 (Component)  : FB_DL_HeaterBreakDetect
 * 所属子库 (Sublibrary) : DL_Device
 * 当前版本 (Version)    : 1.0.0
 * 兼容性   (Platform)   : CODESYS 3.5+ / TwinCAT 3 / 汇川 InoProShop / 施耐德 Machine Expert
 *                         仅依赖 Standard.library（TON / R_TRIG），零厂商私有库
 * 功能描述 (Function)   : 加热管断棒检测（电 + 温双判据，判据介入次序纪律固化）：
 *                         ① 判据一（电流对比）：通电 tWatch 窗到后，电流对基线 fCurRefA 的
 *                            欠偏百分比超 fCurDevPct → eCurLow（电流显著低，直接判低）。
 *                         ② 判据二（温升速率）：**仅在判据一存疑时介入**（电流欠偏为正但
 *                            未达阈值，散热类误报高发域）；以 tTempWatch 自复位窗做窗端温升
 *                            差值判据：窗内温升 < fTempRiseMin × 窗长(分钟) → eNoTempRise。
 *                         ③ 两判据同时成立 → eBreakConfirm **锁存**（断棒确认需人工核查，
 *                            解除沿 = bReset 上升沿）。
 *                         SCR 调功类供电（bPhaseAngle=TRUE，电流与功率非线性）：判据一自动
 *                         降级不判，只信判据二。
 * 接口     (Interface)  : 输入 bHeaterOn 通电、fCurrentA 电流（A）、fTempC 被加热体温度
 *                         （℃）、fCurRefA 额定电流基线（A）、fCurDevPct 判据一欠偏阈值
 *                         （%）、fTempRiseMin 判据二最小温升（℃/min）、tWatch 判据一窗、
 *                         tTempWatch 判据二窗、bPhaseAngle 相角调功声明、bReset 复位；
 *                         输出 eHeat 状态、bError 故障标志。
 * 边界     (Boundary)   : ① **属主边界（写死）：本件只做断棒诊断，不驱动加热器、不调功、
 *                         不接管 SSR/SCR**（驱动归 `FB_DL_SsrHeaterDrive` 族）。
 *                         ② 非通电相全判据冻结回 eOff；温升判据采用窗端差值法（温升 =
 *                         窗末温 - 窗首温），阈值 = fTempRiseMin × 窗长分钟数，分母时间闸
 *                         以窗长 > T#0S 组态闸实现（不做逐拍速率除法，无除零路径）。
 *                         ③ 非有限输入当拍剔除（判据冻结当拍，R245）；窗首温度快照仅在
 *                         有限拍更新（防 NaN 污染快照）。
 *                         ④ TIME_TO_DINT 取窗长毫秒数（tTempWatch 经组态闸保证为正，
 *                         无 TIME_TO_DINT 负值恒假陷阱）。
 *                         ⑤ 组态闸：fCurRefA<=0、fCurDevPct<=0、fTempRiseMin<0、
 *                         tWatch<=T#0S、tTempWatch<=T#0S → 锁存 bError，eHeat 冻结 eOff，
 *                         解除沿 = bReset 上升沿。
 *                         ⑥ 零全局耦合（无 GVL / 无 VAR_EXTERNAL / 无物理地址）。
 * 分工声明 (Scope)      : 与 `FB_DL_SsrHeaterDrive` / `FB_DL_HeaterSsrBank` 分工：诊断
 *                         （本件）≠ 驱动/组 bank（那两件）。
 * 来源标签 (Source Tag) : T2-6 ◐（Rockwell AOI 设备诊断粒度只借"断棒电+温双判据"分类
 *                         事实，判据介入次序纪律为本件自研固化）
 * 码表     (Codes)      : 本件不占用任何全局数字码位。出口为 ENUM 状态 + BOOL；
 *                         数字码位待主控收口阶段统一派号。
 * 红线自检 (Redline)    : R1 ✓ 零 GVL/VAR_EXTERNAL ｜ R2 ✓ 零 %I/%Q/%M ｜ R3 ✓ 纯 IEC 61131-3
 *                         R4 ✓ 除零前置（基线闸）+ 非有限剔除 + 时间域组态闸 ｜ R5 ✓ 声明逐行同行双语注释
 *                         R6 ✓ ENUM 状态判序 ｜ R7 ✓ 两 TON/两 R_TRIG 段 0 无条件刷新
 * 修订历史 (Revision)   : 2026-11-20  v1.0.0  R48 首版（批次 3 · 序号 11）
 *                         验收向量：电流欠偏超阈值 → eCurLow；电流略低 + 窗温升不足 →
 *                         eBreakConfirm 锁存；bPhaseAngle=TRUE 只走温判据；断电回 eOff。
 *==============================================================================*)

TYPE E_DL_HbdState :
(
    eOk           := 0,    // 正常（判据未触发）/ Healthy, no judge fired
    eCurLow       := 10,   // 电流显著欠偏（判据一直接判低）/ Current notably low, judge 1 direct
    eNoTempRise   := 20,   // 温升不足（判据二介入判出）/ Insufficient temperature rise, judge 2 fired
    eBreakConfirm := 30,   // 双判据同时成立，断棒确认（锁存待复位）/ Both judges fired, break confirmed, latched
    eOff          := 40    // 未通电（判据冻结）/ Heater off, judges frozen
);
END_TYPE

FUNCTION_BLOCK FB_DL_HeaterBreakDetect
VAR_INPUT
    bHeaterOn   : BOOL := FALSE;   // 加热器通电状态 [-] / Heater energized state
    fCurrentA   : LREAL := 0.0;    // 加热回路电流实测 [A] / Heater loop current [A]
    fTempC      : LREAL := 0.0;    // 被加热体温度实测 [℃] / Heated body temperature [degC]
    fCurRefA    : LREAL := 10.0;   // 额定电流基线，域 > 0 [A] / Rated current baseline [A]
    fCurDevPct  : LREAL := 30.0;   // 判据一欠偏阈值，域 > 0 [%] / Judge-1 under-deviation threshold [%]
    fTempRiseMin: LREAL := 2.0;    // 判据二最小温升速率，域 >= 0 [℃/min] / Judge-2 minimum rise rate [degC/min]
    tWatch      : TIME := T#10S;   // 判据一观察窗，域 > T#0S [ms] / Judge-1 watch window [ms]
    tTempWatch  : TIME := T#60S;   // 判据二温升窗，域 > T#0S [ms] / Judge-2 rise window [ms]
    bPhaseAngle : BOOL := FALSE;   // 相角调功声明（TRUE=判据一降级只信判据二） [-] / Phase-angle supply declaration
    bReset      : BOOL := FALSE;   // 复位，上升沿清 bError 与断棒锁存 [-] / Reset, rising edge clears latches
END_VAR
VAR_OUTPUT
    eHeat  : E_DL_HbdState;        // 断棒诊断状态出口 [-] / Break-detect state outlet
    bError : BOOL;                 // 故障标志（组态非法 ∨ 断棒确认，锁存） [-] / Error flag, latched
END_VAR
VAR
    _eHeat     : E_DL_HbdState := E_DL_HbdState.eOff;   // 内部状态 / Internal state
    _bCurLow   : BOOL;           // 判据一命中当拍量 / Judge-1 fired this scan
    _bSuspect  : BOOL;           // 判据一存疑（欠偏为正未达阈值）/ Judge-1 suspect flag
    _bNoRise   : BOOL;           // 判据二命中锁存（窗到裁决结果保持到下次裁决）/ Judge-2 fired latch
    _bBreak    : BOOL;           // 断棒确认锁存位（解除沿 = bReset 上升沿） / Break-confirm latch, cleared by reset edge
    _bErrLatch : BOOL;           // 组态故障锁存位（解除沿 = bReset 上升沿） / Latched config fault
    _fTempStart: LREAL := 0.0;   // 温升窗首温度快照 [℃] / Window-start temperature snapshot
    _fRiseLim  : LREAL;          // 温升判据绝对限（速率×窗长分钟） [℃] / Rise judge absolute limit
    _fMinWin   : LREAL;          // 窗长分钟数（毫秒/60000） [min] / Window length in minutes
    _fDevPct   : LREAL;          // 当拍电流欠偏百分比 [%] / Current under-deviation percent
    _bNonFin   : BOOL;           // 输入非有限当拍量 [-] / Non-finite input this scan
    tonWatch   : TON;            // 判据一观察窗定时器，段 0 无条件调用 / Judge-1 window timer
    tonTempWatch: TON;           // 判据二自复位温升窗，段 0 无条件调用 / Judge-2 self-reset rise window
    rtOn       : R_TRIG;         // 通电上升沿实例，段 0 无条件调用 / Energize rising edge instance
    rtReset    : R_TRIG;         // 复位沿实例，段 0 无条件调用 / Reset edge instance
END_VAR
VAR CONSTANT
    DL_HBD_PCT  : LREAL := 100.0;   // 百分比换算基 [无量纲] / Percent conversion base
    DL_HBD_MS   : LREAL := 60000.0; // 毫秒到分钟换算基 [ms/min] / Millisecond-per-minute base
    DL_HBD_ZERO : LREAL := 0.0;     // 非有限差值判零基准 [-] / Non-finite difference zero base
END_VAR

(* —— 段 0：非有限判 + 组态闸 + 两 TON 两沿无条件周期刷新 —— *)
_bNonFin := (fCurrentA <> fCurrentA) OR ((fCurrentA - fCurrentA) <> DL_HBD_ZERO)
         OR (fTempC <> fTempC) OR ((fTempC - fTempC) <> DL_HBD_ZERO);   // 电流/温度非有限（R245） / Non-finite current and temperature
IF (fCurRefA <= 0.0) OR (fCurDevPct <= 0.0) OR (fTempRiseMin < 0.0)
   OR (tWatch <= T#0S) OR (tTempWatch <= T#0S) THEN
    _bErrLatch := TRUE;                                     // 组态域闸：锁存（R188 解除沿 = bReset 上升沿） / Config gate: latch
END_IF
_fMinWin := DINT_TO_LREAL(TIME_TO_DINT(tTempWatch)) / DL_HBD_MS;   // 窗长分钟数（窗长已过正闸，无负值陷阱） / Window minutes
_fRiseLim := fTempRiseMin * _fMinWin;                       // 温升判据绝对限 [℃] / Rise absolute limit
tonWatch(IN := bHeaterOn AND (NOT _bNonFin) AND (NOT _bErrLatch), PT := tWatch);   // 判据一观察窗 / Judge-1 window
tonTempWatch(IN := bHeaterOn AND (NOT tonTempWatch.Q) AND (NOT _bNonFin) AND (NOT _bErrLatch), PT := tTempWatch);   // 判据二自复位窗（R188） / Judge-2 self-reset window
rtOn(CLK := bHeaterOn);                                     // 通电沿，每拍必调 / Energize edge, every scan
rtReset(CLK := bReset);                                     // 复位沿，每拍必调 / Reset edge, every scan

(* —— 段 1：复位沿 / 通电沿（快照初始化） —— *)
IF rtReset.Q THEN
    _bErrLatch := FALSE;                                    // 清组态故障锁存 / Clear config latch
    _bBreak := FALSE;                                       // 清断棒确认锁存 / Clear break latch
    _bNoRise := FALSE;                                      // 清温升判据锁存 / Clear rise latch
END_IF
IF rtOn.Q THEN
    _fTempStart := fTempC;                                  // 通电首拍初始化窗首快照（仅有限拍更新） / Init snapshot on energize
END_IF

(* —— 段 2：判据一（电流对比；相角调功降级不判） —— *)
_bCurLow := FALSE;                                          // 判据一当拍量预清 / Judge-1 preset
_bSuspect := FALSE;                                         // 存疑量预清 / Suspect preset
IF bHeaterOn AND (NOT _bErrLatch) AND (NOT _bNonFin) THEN
    _fDevPct := (fCurRefA - fCurrentA) / fCurRefA * DL_HBD_PCT;   // 欠偏百分比（分母基线已过闸，无除零） / Under-deviation percent
    IF (NOT bPhaseAngle) AND tonWatch.Q THEN
        IF _fDevPct > fCurDevPct THEN
            _bCurLow := TRUE;                               // 判据一直接判低 / Judge-1 direct low
        ELSIF _fDevPct > 0.0 THEN
            _bSuspect := TRUE;                              // 电流略低未达阈值：判据一存疑，判据二获准介入 / Marginally low: judge 2 engaged
        END_IF
    END_IF
END_IF

(* —— 段 3：判据二（窗端温升差值；仅存疑时介入，窗到裁决） —— *)
IF tonTempWatch.Q THEN
    IF _bSuspect AND (NOT _bNonFin) AND ((fTempC - _fTempStart) < _fRiseLim) THEN
        _bNoRise := TRUE;                                   // 窗内温升不足限值：判据二命中（锁存至下次裁决） / Insufficient rise: judge 2 fired
    ELSE
        _bNoRise := FALSE;                                  // 温升达标或无存疑前提：判据二复位 / Rise adequate: judge 2 reset
    END_IF
    _fTempStart := fTempC;                                  // 窗末重置快照（先裁决后重置，防同拍抹除） / Reset snapshot after judging
END_IF

(* —— 段 4：状态合成（断棒确认锁存优先；非通电回 eOff） —— *)
IF _bErrLatch THEN
    _eHeat := E_DL_HbdState.eOff;                           // 组态故障期冻结 eOff 安全侧 / Frozen to eOff on fault
ELSIF NOT bHeaterOn THEN
    _eHeat := E_DL_HbdState.eOff;                           // 非通电相判据冻结 / Off phase frozen
ELSIF _bBreak THEN
    _eHeat := E_DL_HbdState.eBreakConfirm;                  // 锁存回放确认态（不按当下输入重推断，R189） / Latched confirm replay
ELSE
    IF _bCurLow AND _bNoRise THEN
        _bBreak := TRUE;                                    // 双判据同时成立：锁存确认（解除沿 = bReset 上升沿） / Both judges: latch confirm
        _eHeat := E_DL_HbdState.eBreakConfirm;              // 入确认态 / Enter confirm
    ELSIF _bCurLow THEN
        _eHeat := E_DL_HbdState.eCurLow;                    // 判据一单独命中 / Judge 1 alone
    ELSIF _bNoRise THEN
        _eHeat := E_DL_HbdState.eNoTempRise;                // 判据二单独命中 / Judge 2 alone
    ELSE
        _eHeat := E_DL_HbdState.eOk;                        // 判据均未触发 / No judge fired
    END_IF
END_IF

(* —— 段 5：出口单点映射（名实双出口同源，R191） —— *)
eHeat  := _eHeat;                                           // 状态出口 / State outlet
bError := _bErrLatch OR _bBreak;                            // 故障标志 = 组态非法 ∨ 断棒确认 / Error = cfg fault or confirm

END_FUNCTION_BLOCK

(* ---- FB_DL_HeaterSsrBank.st ---- *)
(*
  组件名 Component   : FB_DL_HeaterSsrBank
  子库 Sublibrary    : DL_Device
  版本 Version       : 1.0.0
  兼容性 Platform    : CODESYS 3.5 / TwinCAT 3 / 汇川 InoProShop / Machine Expert（仅 Standard.library）
  功能 Function      : SSR 调功器组（多路时间比例调功 + 均衡 + 断偶降级）：
                       1) 分相输出：各路按 (i-1)/路数 错相起始的时间比例调功（占空比
                       比较内部锯齿相位），错相拉开路间电流峰值，降低电网冲击；
                       2) 路间电流均衡：有效路平均电流基准，单路偏差超 fImbalMaxPct
                       → 均衡告警锁存（维护语义）；
                       3) 断偶/断路降级：占空比高于发波下限而电流低于检测阈，持续
                       tBreakTo 确认 → 该路断偶锁存，出口强制关断（单路降级，其余照常）；
                       4) 每路断偶确认用独立 TON 实例（数组实例，段 0 FOR 无条件刷新）。
  边界 Boundary      : ① 本件只出各路 SSR 开关量与诊断，不写物理 IO；
                       ② 占空比域 [0, 100]，域外钳位 + 均衡告警不置 bError（维护级），
                       断偶锁存置 bError（故障级，bReset 上升沿解除）；
                       ③ 相位换算除法前置域闸：路数域 [1, 8]、周期 > 0；
                       ④ 无全局变量引用、无外部变量声明、无物理地址寻址。
  依赖 Depends       : Standard.library（R_TRIG / TON）
  溯源 Origin        : 道莅自研 clean-room（参考 t2-2-lbp 三段分层分类与参数域，
                       零代码行复制）
  码位 Code          : 16#03_3_1（Device 05xx 副带 0531）
  码表 Error codes（Device 故障窗口 0531，本件无信息码，单故障总码 + 成因枚举归因）:
    16#0003_0531 故障级：SSR 组故障总码（任一路断偶锁存 / 组态非法 / 输入非有限），
                 锁存至 bReset 上升沿，归因见 eCause 与 abChBreak 分量
  修订历史 Revision  :
    2026-11-19  v1.0.0  R44 首版（批次 3 · 序号 13）
*)

TYPE E_DL_HsbState :
(
    eIdle  := 0,    // 空闲：未使能，全路关断 / Idle, all channels off
    eRun   := 10,   // 运行：分相发波 + 诊断 / Running, phased firing and diagnostics
    eFault := 90    // 故障：总码锁存 / Fault, latched
);
END_TYPE

TYPE E_DL_HsbCause :
(
    eNone      := 0,  // 无故障成因 / No cause
    eChBreak   := 1,  // 任一路断偶锁存 / Any channel break latched
    eCfgIllegal:= 2,  // 组态非法 / Illegal configuration
    eNonFinite := 3   // 输入非有限 / Non-finite input
);
END_TYPE

FUNCTION_BLOCK FB_DL_HeaterSsrBank
VAR_INPUT
    bEnable    : BOOL;                     // 使能（电平）[-] / Enable
    bReset     : BOOL;                     // 上升沿清故障锁存 [-] / Reset edge
    nChUse     : INT := 4;                 // 有效路数 [路]，域 1..8 / Active channel count
    afDutyPct  : ARRAY[1..8] OF REAL;      // 各路占空比 [%]，域 0..100 / Duty per channel
    afCurrentA : ARRAY[1..8] OF REAL;      // 各路实测电流 [安培] / Current per channel
    fImbalMaxPct: REAL := 20.0;            // 均衡偏差限 [%] / Imbalance limit
    fBreakDetectA: REAL := 0.5;            // 断偶电流检测阈 [安培] / Break detect threshold
    tPhaseCycle: TIME := T#1S;             // 时间比例周期 [毫秒] / Time-proportional cycle
    tBreakTo   : TIME := T#3S;             // 断偶确认窗 [毫秒] / Break confirm window
END_VAR
VAR_OUTPUT
    abSsrOut   : ARRAY[1..8] OF BOOL;      // 各路 SSR 开关量输出 [-] / SSR output per channel
    abChBreak  : ARRAY[1..8] OF BOOL;      // 各路断偶锁存位 [-] / Break latch per channel
    bImbalAlm  : BOOL;                     // 均衡告警锁存位 [-] / Imbalance alarm latch
    nBreakCount: INT;                      // 断偶路数 [路] / Broken channel count
    eState     : E_DL_HsbState;            // 状态出口，段尾单点映射 / State outlet
    eCause     : E_DL_HsbCause;            // 故障成因出口（R190） / Fault cause outlet
    bError     : BOOL;                     // 故障锁存标志 [-] / Fault latch flag
    uErrId     : UDINT;                    // 事件码，0 = 无事件 / Event code
END_VAR
VAR
    rtReset  : R_TRIG;                     // 复位沿实例，段 0 无条件刷新 / Reset edge
    atonBreak: ARRAY[1..8] OF TON;         // 各路断偶确认实例（数组，段 0 无条件刷新）/ Break timers
    _tPhase  : TIME := T#0S;               // 锯齿相位 [毫秒] / Sawtooth phase
    _eState  : E_DL_HsbState := E_DL_HsbState.eIdle;   // 内部相位（CASE 唯一写入目标）/ Internal phase
    _eCause  : E_DL_HsbCause := E_DL_HsbCause.eNone;   // 故障成因锁存（锁存量）/ Latched cause
    _fPhaseMs: REAL;                       // 相位毫秒值 [毫秒] / Phase in milliseconds
    _fWinMs  : REAL;                       // 周期毫秒值 [毫秒] / Cycle in milliseconds
    _fDutyUse: REAL;                       // 单路钳位占空比 [%] / Clamped duty
    _fAvgA   : REAL;                       // 有效路平均电流 [安培] / Average current
    _nAvgCnt : INT;                        // 有效路计数 [路] / Averaged channel count
    _fImbal  : REAL;                       // 单路偏差 [%] / Per channel imbalance
    _nIdx    : INT;                        // 路索引 [-] / Channel index
    _bFault  : BOOL;                       // 故障锁存位（锁存量） / Latched fault bit
    _uFault  : UDINT;                      // 故障码锁存（锁存量） / Latched fault code
    _bCfgBad : BOOL;                       // 组态非法当拍量 [-] / Config illegal flag
    _bNonFin : BOOL;                       // 输入非有限当拍量 [-] / Non-finite input flag
    _bImbal  : BOOL;                       // 均衡越限当拍量 [-] / Imbalance breach flag
END_VAR
VAR CONSTANT
    DL_CH_MAX   : INT  := 8;               // 路数上限，与数组维度一致 [路] / Channel ceiling
    DL_CH_MIN   : INT  := 1;               // 路数下限 [路] / Channel floor
    DL_DUTY_MAX : REAL := 100.0;           // 占空比上限 [%] / Duty ceiling
    DL_DUTY_MIN : REAL := 0.0;             // 占空比下限 [%] / Duty floor
    DL_DUTY_ONMIN: REAL := 10.0;           // 断偶判据发波下限 [%] / Duty floor for break test
    DL_100      : REAL := 100.0;           // 百分比换算系数 [无量纲] / Percent scale
    DL_ZERO     : REAL := 0.0;             // 零常量 [工程单位] / Zero constant
    DL_ABS_MAX  : REAL := 1.0E30;          // 有限值判定上界 [工程单位] / Finite bound
END_VAR

(* —— 段 0｜沿、相位与定时器每拍无条件刷新（数组实例 FOR 全量刷新，禁置于 CASE 内） —— *)
rtReset(CLK := bReset);
_tPhase := _tPhase + tPhaseCycle;        // 锯齿相位累加（周期性推进）
IF _tPhase >= tPhaseCycle THEN
    _tPhase := _tPhase - tPhaseCycle;    // 相位回卷（差值比较，非取模）
END_IF
_fPhaseMs := TIME_TO_REAL(_tPhase);
_fWinMs   := TIME_TO_REAL(tPhaseCycle);
FOR _nIdx := DL_CH_MIN TO DL_CH_MAX DO
    atonBreak[_nIdx](IN := (_eState = E_DL_HsbState.eRun) AND (NOT _bFault)
                     AND (afDutyPct[_nIdx] >= DL_DUTY_ONMIN)
                     AND (afCurrentA[_nIdx] < fBreakDetectA), PT := tBreakTo);
END_FOR

(* —— 段 1｜瞬时量预清零（锁存量 _bFault/_uFault/abChBreak/bImbalAlm 不入清单） —— *)
uErrId   := 16#0000_0000;
_bCfgBad := FALSE;
_bNonFin := FALSE;
_bImbal  := FALSE;
nBreakCount := 0;
_fAvgA   := DL_ZERO;
_nAvgCnt := 0;

(* —— 段 2｜复位沿：故障与全路断偶锁存一次性清干净（唯一解除路径 = rtReset.Q，
        输入引脚当拍量，调用方拉上升沿即可达） —— *)
IF rtReset.Q THEN
    _bFault := FALSE;
    _uFault := 16#0000_0000;
    _eCause := E_DL_HsbCause.eNone;
    bImbalAlm := FALSE;
    FOR _nIdx := DL_CH_MIN TO DL_CH_MAX DO
        abChBreak[_nIdx] := FALSE;
    END_FOR
    _eState := E_DL_HsbState.eIdle;
END_IF

(* —— 段 3｜组态闸与非有限判据（覆盖全部参与判据换算引脚） —— *)
IF (nChUse < DL_CH_MIN) OR (nChUse > DL_CH_MAX) OR (tPhaseCycle = T#0S)
   OR (fImbalMaxPct <= DL_ZERO) OR (fBreakDetectA <= DL_ZERO) OR (tBreakTo = T#0S) THEN
    _bCfgBad := TRUE;
END_IF
FOR _nIdx := DL_CH_MIN TO DL_CH_MAX DO
    IF (afDutyPct[_nIdx] <> afDutyPct[_nIdx]) OR ((afDutyPct[_nIdx] - afDutyPct[_nIdx]) <> DL_ZERO)
       OR (afCurrentA[_nIdx] <> afCurrentA[_nIdx]) OR ((afCurrentA[_nIdx] - afCurrentA[_nIdx]) <> DL_ZERO) THEN
        _bNonFin := TRUE;
    END_IF
END_FOR

(* —— 段 4｜主状态机：三态全覆盖 + ELSE 兜底 —— *)
CASE _eState OF

E_DL_HsbState.eIdle:
    FOR _nIdx := DL_CH_MIN TO DL_CH_MAX DO
        abSsrOut[_nIdx] := FALSE;        // 空闲相全路关断（安全侧）
    END_FOR
    IF bEnable AND (NOT _bCfgBad) THEN
        _eState := E_DL_HsbState.eRun;
    ELSIF bEnable AND _bCfgBad THEN
        _bFault := TRUE;
        _uFault := 16#0003_0531;
        _eCause := E_DL_HsbCause.eCfgIllegal;
        bError  := TRUE;
        _eState := E_DL_HsbState.eFault;
    END_IF

E_DL_HsbState.eRun:
    IF NOT bEnable THEN
        _eState := E_DL_HsbState.eIdle;  // 使能撤销回空闲
    ELSE
        (* 有效路平均电流基准（仅统计未断偶路） *)
        FOR _nIdx := DL_CH_MIN TO nChUse DO
            IF NOT abChBreak[_nIdx] THEN
                _fAvgA := _fAvgA + afCurrentA[_nIdx];
                _nAvgCnt := _nAvgCnt + 1;
            END_IF
        END_FOR
        IF _nAvgCnt > 0 THEN
            _fAvgA := _fAvgA / INT_TO_REAL(_nAvgCnt);
        END_IF
        FOR _nIdx := DL_CH_MIN TO DL_CH_MAX DO
            IF _nIdx <= nChUse THEN
                (* 分相时间比例调功：窗口起点 = 相位偏移 (i-1)/路数 × 周期 *)
                _fDutyUse := MIN(MAX(afDutyPct[_nIdx], DL_DUTY_MIN), DL_DUTY_MAX);
                IF NOT abChBreak[_nIdx] THEN
                    abSsrOut[_nIdx] := (_fPhaseMs >= (_fWinMs * INT_TO_REAL(_nIdx - 1) / INT_TO_REAL(nChUse)))
                                       AND (_fPhaseMs < (_fWinMs * INT_TO_REAL(_nIdx - 1) / INT_TO_REAL(nChUse)
                                            + _fWinMs * _fDutyUse / DL_100));
                ELSE
                    abSsrOut[_nIdx] := FALSE;    // 断偶路降级强制关断
                END_IF
                (* 断偶确认：Q 置锁存并配对故障码（R45） *)
                IF atonBreak[_nIdx].Q THEN
                    abChBreak[_nIdx] := TRUE;
                    _bFault := TRUE;
                    _uFault := 16#0003_0531;
                    _eCause := E_DL_HsbCause.eChBreak;
                    bError  := TRUE;
                END_IF
            ELSE
                abSsrOut[_nIdx] := FALSE;    // 超出有效路数：强制关断
            END_IF
        END_FOR
        IF _bNonFin THEN
            _bFault := TRUE;                 // 输入非有限：锁存
            _uFault := 16#0003_0531;
            _eCause := E_DL_HsbCause.eNonFinite;
            bError  := TRUE;
            _eState := E_DL_HsbState.eFault;
        ELSE
            (* 均衡监督：有效路偏差超限置告警锁存（维护级，不置 bError） *)
            FOR _nIdx := DL_CH_MIN TO nChUse DO
                IF (NOT abChBreak[_nIdx]) AND (_fAvgA > DL_ZERO) THEN
                    _fImbal := ABS(afCurrentA[_nIdx] - _fAvgA) / _fAvgA * DL_100;
                    IF _fImbal > fImbalMaxPct THEN
                        _bImbal := TRUE;
                    END_IF
                END_IF
            END_FOR
            IF _bImbal THEN
                bImbalAlm := TRUE;           // 均衡告警锁存（bReset 沿解除）
            END_IF
            IF _bFault THEN
                _eState := E_DL_HsbState.eFault;   // 断偶或非有限：进故障相
            END_IF
        END_IF
    END_IF

E_DL_HsbState.eFault:
    FOR _nIdx := DL_CH_MIN TO DL_CH_MAX DO
        abSsrOut[_nIdx] := FALSE;        // 故障相全路关断（安全侧）
    END_FOR
    bError := TRUE;
    ;                                    // 故障相驻留：断偶锁存回放，只认复位沿（段 2 迁出）

ELSE
    _bFault := TRUE;                     // 兜底：非法相位锁存
    _uFault := 16#0003_0531;
    _eCause := E_DL_HsbCause.eCfgIllegal;
    bError  := TRUE;
    _eState := E_DL_HsbState.eFault;
END_CASE

(* —— 段 5｜状态出口单点映射（名实同源） —— *)
eState := _eState;
END_FUNCTION_BLOCK

(* ---- FB_DL_HeatPumpDefrost.st ---- *)
//==============================================================================
// 功能块：FB_DL_HeatPumpDefrost ｜ 中文名称：空气源热泵除霜判据与除霜态时序
// 所属子库：DL_Device ｜ 版本：v1.0.0 ｜ 兼容：CODESYS V3.5+ / TwinCAT 3 / 汇川 InoProShop
// 功能描述：进入三条件：盘管-环境温差达门槛（环境温减盘管温大于等于
//           fCoilAmbDeltaK）、压缩机连续运行达 tMinCompRun、环境温度
//           处于窗口内且湿度达门限；退出：盘管温升至 fExitCoilC 或除
//           霜超时（tDefrostMax）；最小间隔 tDefrostGap 防频繁除霜；
//           超时连续累计供检修判据（MANUAL 建议连续 3 次检修，本件不
//           锁故障：锁死会使机组彻底停机，现场代价高于结霜）。安全侧
//           铁律：任何异常退出都回制热（除霜卡死会让蒸发器彻底结冰）。
//           本件只出请求与状态，四通阀/风机执行由上位裁决。
// 开源溯源 (Origin)：道莅原创实现（参考 公开工程惯例 分类与参数域）
// 单位表：温度[摄氏度] / 温差[K] / 相对湿度[%] / 时长参数[min] / 计数[次]
// 错误码表：16#0003_0192 信息级（除霜请求被最小间隔阻延，阻延沿发一次，
//           不置 bError）/ 16#0003_0193 信息级（除霜超时强制退出回制
//           热，计数累计，不置 bError）/ 16#0003_036C 故障级（参数组
//           态非法，含环境窗倒置、温差门槛非正、任一时长非正、湿度门
//           限超 0~100 域，置 bError）/ 16#0003_036D 故障级（输入非有
//           限，置 bError，强制退出回制热）/ 16#0003_036E 故障级兜底
//           （状态机落 ELSE 或非法状态，置 bError 并强制退出回制热）
// 状态机：E_DL_DefrostState（eIdle=0 / eMonitor=10 / eGapWait=20 /
//           eDefrost=30 / eFault=99），CASE 含 ELSE 兜底，ELSE 置 036E
//           并强制退出除霜回制热（安全侧：除霜态绝不残留）
// 边界行为：① 除霜超时 → 信息 0193 + 强制退出回制热 + uTimeoutCount
//           饱和累计（连续 3 次由 MANUAL 建议检修，不锁故障）；② 环境
//           窗倒置（低大于高）、温差门槛非正、任一时长非正、湿度门限
//           超 0~100 域 → 故障 036C；③ 最小间隔未到 → bBlockedByGap :=
//           TRUE + 信息 0192（请求阻延上升沿发一次，不每拍刷），挂
//           eGapWait，退出条件两条：间隔到（转除霜）或进入条件消失
//           （回监视）；④ 输入非有限（NaN 自反判 + Inf 幅值上限判，
//           R79）→ 故障 036D + 强制退出回制热；⑤ 失能 → 立即退出除
//           霜回制热（安全侧）+ bValid := FALSE；⑥ TON 实例在待机/
//           故障/除霜各分支无条件周期刷新（R40 家族），除霜计时无相
//           内累计；⑦ 首次除霜请求不受间隔约束（上电无历史除霜）；
//           ⑧ 除霜间隔定时器经除霜退出「断输入一拍」重启计时；
//           ⑨ fDeltaK 定义为环境温减盘管温（正值越大结霜趋势越强）。
// 修订历史：v1.0.0 2026-11-17 首版（R25 派单 · §4.5）
//==============================================================================
(*------------------------------------------------------------------------------
 * 枚举: E_DL_DefrostState（归属 DL_Device，与 FB_DL_HeatPumpDefrost 同文件）
 *----------------------------------------------------------------------------*)
TYPE E_DL_DefrostState :
(
    eIdle     := 0,   // 失能/待机：除霜撤、回制热语义 / Idle: defrost withdrawn, back to heating
    eMonitor  := 10,  // 制热监视：三条件逐拍评估 / Monitor: heating, entry conditions evaluated per scan
    eGapWait  := 20,  // 条件满足但最小间隔未到，等待放行 / Conditions met but gap timer running
    eDefrost  := 30,  // 除霜进行中：升温或超时退出 / Defrost active: exits on coil rise or timeout
    eFault    := 99   // 故障兜底态：组态非法/非有限/非法状态，强制回制热 / Fault fallback, forced back to heating
);
END_TYPE
FUNCTION_BLOCK FB_DL_HeatPumpDefrost
VAR_INPUT
    fCoilC        : LREAL;                       // 盘管温度 [摄氏度] / Coil temperature [degC]
    fAmbC         : LREAL;                       // 环境温度 [摄氏度] / Ambient temperature [degC]
    fAmbRhPct     : LREAL;                       // 环境相对湿度 [百分数] / Ambient relative humidity [percent]
    bCompRunning  : BOOL;                        // 压缩机运行反馈 / Compressor running feedback
    fCoilAmbDeltaK : LREAL := 8.0;               // 进入温差门槛 [K]（环境减盘管）/ Entry delta threshold [K], ambient minus coil
    fAmbWinLowC   : LREAL := -5.0;               // 环境温度窗下限 [摄氏度] / Ambient window lower bound [degC]
    fAmbWinHighC  : LREAL := 15.0;               // 环境温度窗上限 [摄氏度] / Ambient window upper bound [degC]
    fRhMinPct     : LREAL := 50.0;               // 湿度门限 [百分数] / Humidity threshold [percent]
    fExitCoilC    : LREAL := 12.0;               // 退出盘管温 [摄氏度] / Exit coil temperature [degC]
    tMinCompRun   : TIME := T#45M;               // 压缩机连续运行门槛 [min] / Minimum continuous compressor run [min]
    tDefrostMax   : TIME := T#10M;               // 除霜最大时长 [min] / Maximum defrost duration [min]
    tDefrostGap   : TIME := T#30M;               // 两次除霜最小间隔 [min] / Minimum interval between defrosts [min]
    bEnable       : BOOL;                        // 总使能 / Master enable
    bReset        : BOOL;                        // 复位，上升沿清状态与计数 / Reset, rising edge clears state and counters
END_VAR
VAR_OUTPUT
    bDefrostReq   : BOOL;                       // 除霜请求（条件满足且未在除霜中）/ Defrost request (conditions met and not active)
    bDefrostActive : BOOL;                      // 除霜进行中 / Defrost active flag
    tDefrostElapsed : TIME;                     // 除霜已进行时长 [min]：除霜中实时，退出后保持末次时长（诊断用）/ Elapsed defrost duration, live while active, holds last value after exit for diagnostics
    fDeltaK       : LREAL;                      // 结霜趋势温差 [K]，环境减盘管 / Frost-trend delta [K], ambient minus coil
    bBlockedByGap : BOOL;                       // 请求被最小间隔阻延 / Request blocked by gap interval
    bOutOfWindow  : BOOL;                       // 环境温度在窗外 / Ambient temperature out of window
    uDefrostCount : UDINT;                      // 累计除霜次数 [次]，饱和计数 / Cumulative defrost count, saturated
    uTimeoutCount : UDINT;                      // 累计除霜超时次数 [次]，饱和计数 / Cumulative timeout count, saturated
    eErr          : UDINT;                      // 错误码，0 = 无错，码位 16#0003_0192 起信息级、16#0003_036C 起故障级（分带见错误码表） / Error code, 0 = no error, band info/fault per the code table
    bError        : BOOL;                       // 故障级标志，仅故障级错误置位 / Fault-class flag, set only on fault-level codes
    bValid        : BOOL;                       // 判据数据可用标志，失能/故障闸显式 FALSE / Verdict usable flag, explicit FALSE on disable/fault gates
    eState        : E_DL_DefrostState;          // 主状态机当前状态 / Current state of the main state machine
END_VAR
VAR
    fbReset       : R_TRIG;                     // 复位上升沿检测实例 / Reset rising edge detector
    fbCompRun     : TON;                        // 压缩机连续运行定时器 / Continuous compressor run timer
    fbDefrost     : TON;                        // 除霜时长定时器（超时判据）/ Defrost duration timer, timeout basis
    fbGap         : TON;                        // 除霜最小间隔定时器 / Defrost gap interval timer
    bGapKick      : BOOL;                       // 间隔定时器断输入一拍标志（R40 家族）/ Gap timer one-scan kick flag
    fbReqBlockTrig : R_TRIG;                    // 请求阻延上升沿检测实例（0192 一次触发）/ Request-block rising edge detector, 0192 once per edge
    bEnterCond    : BOOL;                       // 除霜进入三条件全满足 / All three entry conditions met
    bGapOk        : BOOL;                       // 间隔放行：无历史除霜或间隔已满 / Gap released: no history or interval elapsed
    bBlockedNow   : BOOL;                       // 本拍请求被阻延 / Request blocked this scan
    bDefrostEver  : BOOL;                       // 激活以来是否除过霜 / Any defrost since activation
END_VAR
VAR CONSTANT
    DL_HPD_CODE_INFO_1 : UDINT := 16#0003_0192;   // 信息级槽 1（请求被最小间隔阻延） / info slot 1
    DL_HPD_CODE_INFO_2 : UDINT := 16#0003_0193;   // 信息级槽 2（除霜超时强制退出） / info slot 2
    DL_HPD_CODE_FLT_1  : UDINT := 16#0003_036C;   // 故障级槽 1（参数组态非法） / fault slot 1
    DL_HPD_CODE_FLT_2  : UDINT := 16#0003_036D;   // 故障级槽 2（输入非有限） / fault slot 2
    DL_HPD_CODE_FLT_3  : UDINT := 16#0003_036E;   // 故障级槽 3（非法状态兜底） / fault slot 3, illegal-state fallback
    DL_DF_ZERO    : LREAL := 0.0;               // 零值常量，避免裸字面量 [—] / Zero constant, avoids a bare literal
    DL_DF_TOL     : LREAL := 1.0E-6;            // 浮点比较容差 [—] / Float comparison tolerance
    DL_DF_INF     : LREAL := 1.7976931348623157E308;  // LREAL 幅值上限，Inf 判据 / LREAL magnitude ceiling, Inf criterion
    DL_DF_CNT_MAX : UDINT := 16#FFFF_FFFE;      // 饱和计数上限 [次] / Saturating counter ceiling
    DL_DF_RH_MAX  : LREAL := 100.0;             // 湿度门限域上限 [百分数] / Humidity threshold domain ceiling [percent]
END_VAR

(*------------------------------------------------------------------------------
 * 段 1｜无条件刷新区（红线 5）：三 TON 与两 R_TRIG 在任何分支之外周期调用
 *----------------------------------------------------------------------------*)
fbReset(CLK := bReset);                        // 复位沿检测无条件刷新 / reset edge refreshed unconditionally
fbCompRun(IN := bCompRunning AND bEnable,      // 压缩机连续运行计时（失能即断）/ compressor run timing, broken on disable
          PT := tMinCompRun);                  // 连续运行门槛 / continuous run threshold
fbDefrost(IN := (eState = E_DL_DefrostState.eDefrost) AND bEnable,  // 仅除霜态计时（相内不累计，R40 家族）/ times only in defrost state
          PT := tDefrostMax);                  // 除霜最大时长 / maximum defrost duration
fbGap(IN := bEnable AND NOT bGapKick,          // 间隔计时，断输入一拍重启（R40 家族）/ gap timing, kicked one scan per defrost exit
      PT := tDefrostGap);                      // 最小间隔 / minimum interval
bGapKick := FALSE;                             // kick 标志单拍自清（除霜退出时由状态机重置位）/ kick self-clears, state machine re-sets on exit

(*------------------------------------------------------------------------------
 * 段 2｜复位沿处理（改写置于沿后，防吞沿 R39）
 *----------------------------------------------------------------------------*)
IF fbReset.Q THEN
    eState        := E_DL_DefrostState.eIdle;
    eErr          := 16#0000_0000;             // 复位清码 / reset clears code
    bError        := FALSE;                    // 复位清故障 / reset clears fault
    bDefrostReq   := FALSE;                    // 请求撤 / request withdrawn
    bDefrostActive := FALSE;                   // 除霜撤（回制热语义）/ defrost withdrawn
    bBlockedByGap := FALSE;                    // 阻延标志清 / block flag cleared
    uDefrostCount := 0;                        // 除霜计数清零 / defrost count zeroed
    uTimeoutCount := 0;                        // 超时计数清零 / timeout count zeroed
    bDefrostEver  := FALSE;                    // 除霜历史清零，首个请求放行 / defrost history cleared, first request released
END_IF

(*------------------------------------------------------------------------------
 * 段 3｜非有限输入闸（浮点引脚逐个：NaN 自反判 + Inf 幅值上限判，R79）
 *       命中即强制退出除霜回制热（安全侧）
 *----------------------------------------------------------------------------*)
IF (fCoilC <> fCoilC) OR (ABS(fCoilC) >= DL_DF_INF)
   OR (fAmbC <> fAmbC) OR (ABS(fAmbC) >= DL_DF_INF)
   OR (fAmbRhPct <> fAmbRhPct) OR (ABS(fAmbRhPct) >= DL_DF_INF)
   OR (fCoilAmbDeltaK <> fCoilAmbDeltaK) OR (ABS(fCoilAmbDeltaK) >= DL_DF_INF)
   OR (fAmbWinLowC <> fAmbWinLowC) OR (ABS(fAmbWinLowC) >= DL_DF_INF)
   OR (fAmbWinHighC <> fAmbWinHighC) OR (ABS(fAmbWinHighC) >= DL_DF_INF)
   OR (fRhMinPct <> fRhMinPct) OR (ABS(fRhMinPct) >= DL_DF_INF)
   OR (fExitCoilC <> fExitCoilC) OR (ABS(fExitCoilC) >= DL_DF_INF) THEN
    eState         := E_DL_DefrostState.eFault;
    eErr           := DL_HPD_CODE_FLT_2;           // 故障级：输入非有限 / fault: non-finite input
    bError         := TRUE;                    // 故障级必置 bError（R45 配对）/ fault-class pairs with bError
    bValid         := FALSE;                   // 输出不可用 / outputs unusable
    bDefrostReq    := FALSE;                   // 请求撤 / request withdrawn
    bDefrostActive := FALSE;                   // 强制退出回制热（安全侧）/ forced back to heating, safe side
    bBlockedByGap  := FALSE;                   // 阻延标志清 / block flag cleared
    bOutOfWindow   := FALSE;                   // 故障态不判窗外 / out-of-window not judged in fault
    tDefrostElapsed := fbDefrost.ET;           // 时长出口为定时器实值（已断输入归零）/ elapsed output mirrors timer (input broken, zeroed)
    fbReqBlockTrig(CLK := FALSE);              // 阻延沿检测无条件刷新（早退路径保刷新，红线 5）/ block edge refreshed unconditionally on early-exit path
    RETURN;
END_IF

(*------------------------------------------------------------------------------
 * 段 4｜参数组态闸（窗倒置/温差门槛非正/任一时长非正/湿度门限超域/退出温非正）
 *----------------------------------------------------------------------------*)
IF (fAmbWinLowC > fAmbWinHighC)
   OR (fCoilAmbDeltaK <= DL_DF_TOL)
   OR (tMinCompRun <= T#0S) OR (tDefrostMax <= T#0S) OR (tDefrostGap <= T#0S)
   OR (fRhMinPct < DL_DF_ZERO) OR (fRhMinPct > DL_DF_RH_MAX)
   OR (fExitCoilC <= DL_DF_ZERO) THEN
    eState         := E_DL_DefrostState.eFault;
    eErr           := DL_HPD_CODE_FLT_1;           // 故障级：参数组态非法 / fault: parameter config invalid
    bError         := TRUE;                    // 故障级必置 bError（R45 配对）/ fault-class pairs with bError
    bValid         := FALSE;                   // 输出不可用 / outputs unusable
    bDefrostReq    := FALSE;                   // 请求撤 / request withdrawn
    bDefrostActive := FALSE;                   // 强制退出回制热（安全侧）/ forced back to heating, safe side
    bBlockedByGap  := FALSE;                   // 阻延标志清 / block flag cleared
    bOutOfWindow   := FALSE;                   // 故障态不判窗外 / out-of-window not judged in fault
    tDefrostElapsed := fbDefrost.ET;           // 时长出口为定时器实值 / elapsed output mirrors timer
    fbReqBlockTrig(CLK := FALSE);              // 阻延沿检测无条件刷新（早退路径保刷新，红线 5）/ block edge refreshed unconditionally on early-exit path
    RETURN;
END_IF

(*------------------------------------------------------------------------------
 * 段 5｜判据计算：温差、窗外、进入三条件、间隔放行、阻延
 *----------------------------------------------------------------------------*)
fDeltaK := fAmbC - fCoilC;                     // 结霜趋势温差 = 环境 − 盘管 [K] / frost-trend delta [K]
bOutOfWindow := (fAmbC < fAmbWinLowC) OR (fAmbC > fAmbWinHighC);  // 环境窗外 / ambient out of window
bEnterCond := (fDeltaK >= fCoilAmbDeltaK)      // 条件一：温差达门槛 / condition 1: delta threshold
          AND fbCompRun.Q                     // 条件二：压缩机连续运行达门槛 / condition 2: continuous run
          AND (NOT bOutOfWindow)              // 条件三之一：环境在窗内 / condition 3a: in window
          AND (fAmbRhPct >= fRhMinPct)        // 条件三之二：湿度达门限 / condition 3b: humidity threshold
          AND bCompRunning;                   // 压缩机运行中（除霜只在运行态进）/ compressor running
bGapOk := (NOT bDefrostEver) OR fbGap.Q;       // 间隔放行：无历史除霜或最小间隔已满 / gap released
bBlockedNow := bEnterCond AND (NOT bGapOk);    // 本拍阻延判据 / blocked predicate this scan
fbReqBlockTrig(CLK := bBlockedNow);            // 阻延沿检测无条件刷新（0192 沿发一次）/ block edge refreshed unconditionally

(*------------------------------------------------------------------------------
 * 段 6｜状态机：CASE 含 ELSE 兜底（非法状态 → 036E + 强制回制热，安全侧）
 *----------------------------------------------------------------------------*)
bDefrostActive := (eState = E_DL_DefrostState.eDefrost);  // 除霜态先行取值（CASE 改写前）/ defrost flag captured before CASE rewrite

CASE eState OF

    E_DL_DefrostState.eIdle:
        bValid := FALSE;                       // 失能闸显式不可用（R72）/ explicit FALSE on disable gate
        bDefrostReq := FALSE;                  // 请求撤 / request withdrawn
        bDefrostActive := FALSE;               // 除霜撤（回制热语义）/ defrost withdrawn
        bBlockedByGap := FALSE;                // 阻延标志清 / block flag cleared
        eErr := 16#0000_0000;                  // 待机无错 / no error in idle
        bError := FALSE;                       // 待机无故障 / no fault in idle
        IF bEnable THEN
            eState := E_DL_DefrostState.eMonitor;      // 使能进制热监视 / enable enters heating monitor
        END_IF

    E_DL_DefrostState.eMonitor:
        bValid := TRUE;                        // 监视态判据可用 / verdict usable in monitor
        bDefrostActive := FALSE;               // 非除霜态 / not defrosting
        bDefrostReq := bEnterCond AND (NOT bGapOk);  // 请求被阻延时仍如实外显 / request shown while blocked
        bBlockedByGap := bBlockedNow;          // 阻延标志逐拍刷新 / block flag refreshed per scan
        IF bEnterCond AND bGapOk THEN
            eState := E_DL_DefrostState.eDefrost;      // 三条件齐且间隔放行：进除霜 / conditions met and gap released: defrost
            bDefrostEver := TRUE;              // 记录除霜历史 / record defrost history
            uDefrostCount := uDefrostCount + 1;        // 除霜计数累计 / defrost count up
            IF uDefrostCount >= DL_DF_CNT_MAX THEN
                uDefrostCount := DL_DF_CNT_MAX;        // 饱和防回绕 / saturate to avoid wrap
            END_IF
        ELSIF bEnterCond THEN
            eState := E_DL_DefrostState.eGapWait;      // 条件齐但间隔未到：挂起等待 / conditions met but gap running: wait
        END_IF

    E_DL_DefrostState.eGapWait:
        bValid := TRUE;                        // 等待态判据可用 / verdict usable in wait
        bDefrostActive := FALSE;               // 非除霜态 / not defrosting
        bDefrostReq := TRUE;                   // 请求保持外显 / request held visible
        bBlockedByGap := TRUE;                 // 阻延标志保持 / block flag held
        IF NOT bEnable THEN
            eState := E_DL_DefrostState.eIdle;         // 失能回待机（安全侧）/ disable returns to idle
            bValid := FALSE;                   // 失能闸显式不可用 / explicit FALSE on disable gate
            bDefrostReq := FALSE;              // 请求撤 / request withdrawn
            bBlockedByGap := FALSE;            // 阻延标志清 / block flag cleared
        ELSIF NOT bEnterCond THEN
            eState := E_DL_DefrostState.eMonitor;      // 进入条件消失退出（第二条退出条件）/ entry conditions vanished, second exit
            bDefrostReq := FALSE;              // 请求撤 / request withdrawn
            bBlockedByGap := FALSE;            // 阻延标志清 / block flag cleared
        ELSIF fbGap.Q THEN
            eState := E_DL_DefrostState.eDefrost;      // 间隔到转除霜（第一条退出条件）/ gap elapsed, first exit: defrost
            bDefrostEver := TRUE;              // 记录除霜历史 / record defrost history
            uDefrostCount := uDefrostCount + 1;        // 除霜计数累计 / defrost count up
            IF uDefrostCount >= DL_DF_CNT_MAX THEN
                uDefrostCount := DL_DF_CNT_MAX;        // 饱和防回绕 / saturate to avoid wrap
            END_IF
        END_IF

    E_DL_DefrostState.eDefrost:
        bValid := TRUE;                        // 除霜态判据可用 / verdict usable in defrost
        bDefrostActive := TRUE;                // 除霜进行中 / defrosting
        bDefrostReq := FALSE;                  // 已在除霜，请求撤 / already defrosting, request withdrawn
        bBlockedByGap := FALSE;                // 除霜中无阻延语义 / no blocking semantics in defrost
        tDefrostElapsed := fbDefrost.ET;       // 除霜时长出口 [min] / elapsed defrost duration
        IF fCoilC >= fExitCoilC THEN
            eState := E_DL_DefrostState.eMonitor;      // 盘管升温正常退出 / coil warmed, normal exit
            bGapKick := TRUE;                  // 间隔定时器断输入一拍重启 / gap timer kicked one scan
            bDefrostActive := FALSE;           // 回制热（安全侧）/ back to heating, safe side
        ELSIF fbDefrost.Q THEN
            eState := E_DL_DefrostState.eMonitor;      // 超时强制退出回制热（安全侧）/ timeout forced exit back to heating
            eErr := DL_HPD_CODE_INFO_2;        // 信息级：除霜超时强制退出 / info: defrost timeout forced exit
            bError := FALSE;                   // 信息级不置 bError / info never raises bError
            uTimeoutCount := uTimeoutCount + 1;        // 超时计数累计（检修判据）/ timeout count up, maintenance evidence
            IF uTimeoutCount >= DL_DF_CNT_MAX THEN
                uTimeoutCount := DL_DF_CNT_MAX;        // 饱和防回绕 / saturate to avoid wrap
            END_IF
            bGapKick := TRUE;                  // 间隔定时器断输入一拍重启 / gap timer kicked one scan
            bDefrostActive := FALSE;           // 回制热（安全侧）/ back to heating, safe side
        END_IF

    ELSE
        eState := E_DL_DefrostState.eFault;    // 非法状态兜底 / illegal-state fallback
        eErr := DL_HPD_CODE_FLT_3;                 // 故障级兜底：非法状态 / fault fallback: illegal state
        bError := TRUE;                        // 故障级必置 bError / fault-class pairs with bError
        bValid := FALSE;                       // 输出不可用 / outputs unusable
        bDefrostReq := FALSE;                  // 请求撤 / request withdrawn
        bDefrostActive := FALSE;               // 强制退出回制热（安全侧，除霜态绝不残留）/ forced back to heating, never residual
        bBlockedByGap := FALSE;                // 阻延标志清 / block flag cleared
END_CASE

(*------------------------------------------------------------------------------
 * 段 7｜信息级收口：阻延沿发一次 0192（不每拍刷，见边界行为③）
 *----------------------------------------------------------------------------*)
IF fbReqBlockTrig.Q THEN
    eErr := DL_HPD_CODE_INFO_1;                // 信息级：除霜请求被最小间隔阻延 / info: defrost request blocked by gap
    bError := FALSE;                           // 信息级不置 bError / info never raises bError
END_IF
END_FUNCTION_BLOCK

(* ---- FB_DL_HeatTraceCircuitMon.st ---- *)
(*
  Name        : FB_DL_HeatTraceCircuitMon
  Category    : DL_Device
  Version     : 1.0.1
  Purpose     : 电伴热回路监视：以「加热命令 × 电流存在性 × 温升响应」三重交叉判据区分断缆（无电流）、空烧/过热（超温）、热耦合失效（有电流但无温升）；/ Monitor heat-trace circuits by cross-checking heat command, current presence and temperature-rise response to distinguish open circuit, over-temperature and lost thermal coupling
  溯源        : 借 t2-8-isa182·回路一致性 的分类/参数域组织，clean-room 实现
  Boundary    : ① 组态闸：电流下限/观察窗/最小温升/温度上限任一越域 → 锁存故障；
                ② 观察窗用自复位 TON（IN := NOT tonObs.Q，R188），窗起点温度快照在窗开始那拍取；
                ③ 断缆判据需延时确认（tCurrentConf），避免接触器合闸瞬态误判；
                ④ 三种成因各有独立状态成员与独立判据位（R190 归因唯一），不共用枚举成员；
                ⑤ 本件为诊断层，不驱动加热输出；切除动作须由上层安全联锁执行（属主边界）。
                ⑥ 输出语义（R191 名实双出口）：三个判据位在命中后锁存（仅复位沿清），bError 与
                   之同源置位；相位保持在 eMon 继续监视（不迁 eFault 冻结），以便断缆修复后
                   仍能观察其余判据 —— 此为「降级继续监视」而非冻结，故不置 eFault。
  修订记录    : 2026-11-20 v1.0.1：段 0 双定时器 IN 串 eMon 相位闸（确认延时/观察窗不再跨相自由跑，R52-07）；eIdle→eMon 迁入拍补 _fTempT0/_bT0Ok 起点快照。
*)
TYPE E_DL_HtcState :
(
    eIdle  := 0,                             (* 未使能 / Disabled *)
    eMon   := 10,                            (* 监视运行 / Monitoring *)
    eFault := 90                             (* 故障锁存相 / Fault latched *)
);
END_TYPE

TYPE E_DL_HtcCause :
(
    eNone       := 0,                        (* 无故障成因 / No cause *)
    eCfgIllegal := 1,                        (* 组态非法：电流/时间/温升/温度越域 / Illegal config *)
    eOpenCirc   := 2,                        (* 成因：断缆（命令通而无电流） / Cause: open circuit *)
    eOverTemp   := 3,                        (* 成因：过热（超温上限） / Cause: over-temperature *)
    eNoRise     := 4,                        (* 成因：无温升（电流有而热耦合失效） / Cause: no temperature rise *)
    ePhaseBad   := 5                         (* 非法相位兜底 / Illegal phase fallback *)
);
END_TYPE

FUNCTION_BLOCK FB_DL_HeatTraceCircuitMon
VAR_INPUT
    bHeatCmd   : BOOL := FALSE;              (* 加热命令电平 [-] / Heat command level *)
    fCurrent   : REAL := 0.0;                (* 回路电流实测，域 >= 0 [A] / Measured loop current *)
    fCurrentMin: REAL := 0.5;                (* 电流存在性下限，域 > 0 [A] / Current presence threshold, > 0 *)
    fTemp      : REAL := 20.0;               (* 伴热测点温度 [°C] / Heat-trace temperature *)
    tObserve   : TIME := T#300S;             (* 温升观察窗长，域 > T#0S [ms] / Rise observation window, > 0 *)
    fRiseMin   : REAL := 3.0;                (* 窗内最小期望温升，域 > 0 [K] / Minimum expected rise, > 0 *)
    fTempMax   : REAL := 120.0;              (* 温度上限（过热阈值）[°C] / Over-temperature limit *)
    bEnable    : BOOL := TRUE;               (* 监视使能 [-] / Enable *)
    bReset     : BOOL := FALSE;              (* 复位命令，上升沿清锁存与故障 [-] / Reset command *)
END_VAR
VAR_OUTPUT
    fRiseObs   : REAL;                       (* 观察窗内实测温升（当前窗）[K] / Measured rise in current window *)
    bCurPresent: BOOL;                       (* 电流存在性（本拍判定）[-] / Current presence *)
    bOpenCirc  : BOOL;                       (* 断缆判据锁存（命令通且无电流）[-] / Open-circuit latch *)
    bOverTemp  : BOOL;                       (* 过热判据锁存（超温上限）[-] / Over-temperature latch *)
    bNoRise    : BOOL;                       (* 无温升判据锁存（有电流但窗内温升不足）[-] / No-rise latch *)
    eState     : E_DL_HtcState;              (* 状态出口 / State outlet *)
    eCause     : E_DL_HtcCause;              (* 故障成因出口（R190 归因唯一） / Fault cause outlet *)
    bError     : BOOL;                       (* 故障锁存标志 [-] / Fault latch flag *)
END_VAR
VAR
    _eState  : E_DL_HtcState := E_DL_HtcState.eIdle;     (* 内部相位（CASE 唯一写入目标） / Internal phase *)
    _eCause  : E_DL_HtcCause := E_DL_HtcCause.eNone;     (* 故障成因锁存量 / Latched cause *)
    rtReset  : R_TRIG;                       (* 复位沿实例，段 0 无条件调用 / Reset edge instance *)
    tonObs   : TON;                          (* 观察窗自复位计时器（R188） / Self-resetting observation window *)
    tonNoCur : TON;                          (* 无电流确认延时计时器（IN 由命令与电流派生） / No-current confirm timer *)
    _bFault  : BOOL;                         (* 故障锁存位 / Latched fault bit *)
    _bCfgBad : BOOL;                         (* 组态非法当拍量 / Illegal config this scan *)
    _bFinite : BOOL;                         (* 输入有限性当拍量 / Input finiteness *)
    _bCur    : BOOL;                         (* 电流存在性当拍量 / Current presence this scan *)
    _fTempT0 : REAL;                         (* 观察窗起点温度快照 [°C] / Temperature at window start *)
    _bT0Ok   : BOOL;                         (* 起点快照有效标志 / Snapshot validity *)
    _fRise   : REAL;                         (* 本窗温升中间量 [K] / Rise intermediate *)
END_VAR
VAR CONSTANT
    DL_HTC_EPS    : REAL := 1.0E-6;          (* 判零容差 [-] / Epsilon *)
    DL_HTC_TMIN   : REAL := 0.0;             (* 温度上限可接受下限（防组态倒置）[°C] / Temperature limit floor *)
    DL_HTC_CONF   : TIME := T#5S;            (* 断缆确认延时（接触器合闸瞬态穿越）[ms] / Open-circuit confirm delay *)
END_VAR

(* —— 段 0：当拍判据派生 + 实例无条件刷新（R228A；定时器全在段 0，无 IF 包裹） —— *)
_bCfgBad := (fCurrentMin <= DL_HTC_EPS)                                        (* 电流下限正域闸 / Current threshold gate *)
            OR NOT (tObserve > T#0S)                                           (* 观察窗正域闸 / Window gate *)
            OR (fRiseMin <= DL_HTC_EPS)                                        (* 最小温升正域闸 / Rise gate *)
            OR (fTempMax < DL_HTC_TMIN);                                       (* 温度上限须为非负（防组态倒置） / Temperature limit gate *)
rtReset(CLK := bReset);                                                        (* 复位沿每拍必调 / Reset edge every scan *)
tonObs(IN := (_eState = E_DL_HtcState.eMon) AND NOT tonObs.Q, PT := tObserve);                 (* 观察窗自复位（R188）+ eMon 相位闸（v1.0.1，上拍相位 1 拍延迟可接受） / Self-resetting window with phase gate *)
tonNoCur(IN := (_eState = E_DL_HtcState.eMon) AND bHeatCmd AND NOT _bCur, PT := DL_HTC_CONF);   (* 无电流确认延时（命令通且无电流才计时）+ 相位闸（v1.0.1） / No-current confirm with phase gate *)
_bFinite := (fCurrent = fCurrent) AND (fTemp = fTemp)                          (* NaN 自反闸 / NaN reflex gates *)
            AND ((fCurrent - fCurrent) = (fCurrent - fCurrent))                (* 电流 Inf 闸 / Current Inf gate *)
            AND ((fTemp - fTemp) = (fTemp - fTemp));                           (* 温度 Inf 闸 / Temperature Inf gate *)
_bCur := _bFinite AND (fCurrent >= fCurrentMin);                               (* 电流存在性：有限且 >= 下限 / Presence: finite and above threshold *)

(* —— 段 1：单拍量预清零（R107） —— *)
bCurPresent := FALSE;                                                          (* 电流指示预清 / Presence preset *)
fRiseObs := 0.0;                                                               (* 温升出口预清 / Rise preset *)

(* —— 段 2：复位沿处理（作用域：清故障 + 清三判据 + 清快照 + 迁 eIdle，R283 逐项声明） —— *)
IF rtReset.Q THEN
    _bFault := FALSE;                                                          (* 清故障锁存 / Clear fault *)
    _eCause := E_DL_HtcCause.eNone;                                            (* 清成因 / Clear cause *)
    bOpenCirc := FALSE;                                                        (* 清断缆判据 / Clear open-circuit *)
    bOverTemp := FALSE;                                                        (* 清过热判据 / Clear over-temperature *)
    bNoRise := FALSE;                                                          (* 清无温升判据 / Clear no-rise *)
    _bT0Ok := FALSE;                                                           (* 清起点快照有效位（重新取快照） / Clear snapshot flag *)
    _fTempT0 := 0.0;                                                           (* 清起点温度 / Clear snapshot value *)
    _eState := E_DL_HtcState.eIdle;                                            (* 迁未使能相 / Back to idle *)
END_IF

(* —— 段 3：组态故障锁存（锁存至复位沿，R189） —— *)
IF _bCfgBad AND NOT _bFault THEN
    _bFault := TRUE;                                                           (* 锁存故障位 / Latch fault *)
    _eCause := E_DL_HtcCause.eCfgIllegal;                                      (* 成因：组态非法 / Cause: illegal config *)
    _eState := E_DL_HtcState.eFault;                                           (* 同步迁故障相 / Migrate to fault *)
END_IF

(* —— 段 4：CASE 主状态机（ELSE 兜底迁 eFault，红线 6） —— *)
CASE _eState OF
    E_DL_HtcState.eIdle:                                                       (* 未使能：快照失效，不判 / Disabled *)
        _bT0Ok := FALSE;                                                       (* 失能清快照（重使能重新对齐） / Clear snapshot *)
        IF bEnable AND NOT _bFault THEN
            _fTempT0 := fTemp;                                                 (* 迁入拍即取窗起点温度快照（相位闸配套，v1.0.1） / Snapshot at entry scan *)
            _bT0Ok := TRUE;                                                    (* 快照有效位随迁入同步置位 / Set snapshot flag at entry *)
            _eState := E_DL_HtcState.eMon;                                     (* 使能进入监视 / Enter monitoring *)
        END_IF
    E_DL_HtcState.eMon:                                                        (* 监视相：三重判据 / Monitoring *)
        IF NOT bEnable THEN
            _eState := E_DL_HtcState.eIdle;                                    (* 失能回未使能 / Back to idle *)
        ELSE
            bCurPresent := _bCur;                                              (* 电流指示出口（名实同源，R191） / Presence outlet *)
            IF _bFinite THEN
                IF NOT _bT0Ok THEN
                    _fTempT0 := fTemp;                                         (* 窗起点快照：首拍或窗回零点 / Window start snapshot *)
                    _bT0Ok := TRUE;                                            (* 立快照有效位 / Set snapshot flag *)
                END_IF
                _fRise := fTemp - _fTempT0;                                    (* 本窗温升 = 当前 - 起点（可负）[K] / Rise this window *)
                fRiseObs := _fRise;                                            (* 温升出口 / Rise outlet *)
                IF fTemp > fTempMax THEN                                       (* 过热判据（独立位，R190） / Over-temperature verdict *)
                    bOverTemp := TRUE;                                         (* 过热锁存（复位沿清） / Latch over-temperature *)
                    IF NOT _bFault THEN
                        _bFault := TRUE;                                       (* 同步故障锁存 / Latch fault *)
                        _eCause := E_DL_HtcCause.eOverTemp;                    (* 成因：过热 / Cause: over-temperature *)
                    END_IF
                END_IF
                IF tonNoCur.Q THEN                                             (* 命令通但确认延时内无电流：断缆 / Open circuit *)
                    bOpenCirc := TRUE;                                         (* 断缆锁存（复位沿清） / Latch open-circuit *)
                    IF NOT _bFault THEN
                        _bFault := TRUE;                                       (* 同步故障锁存 / Latch fault *)
                        _eCause := E_DL_HtcCause.eOpenCirc;                    (* 成因：断缆 / Cause: open circuit *)
                    END_IF
                END_IF
                IF tonObs.Q THEN                                               (* 观察窗到点：结算温升响应 / Window elapsed: settle *)
                    IF _bCur AND (_fRise < fRiseMin) THEN                      (* 有电流却温升不足：热耦合失效 / Current present but no rise *)
                        bNoRise := TRUE;                                       (* 无温升锁存（复位沿清） / Latch no-rise *)
                        IF NOT _bFault THEN
                            _bFault := TRUE;                                   (* 同步故障锁存 / Latch fault *)
                            _eCause := E_DL_HtcCause.eNoRise;                  (* 成因：无温升 / Cause: no rise *)
                        END_IF
                    END_IF
                    _fTempT0 := fTemp;                                         (* 新窗起点重置（自复位计时器同拍已回 0） / Restart window baseline *)
                    _bT0Ok := TRUE;                                            (* 快照保持有效 / Keep snapshot valid *)
                END_IF
            END_IF                                                             (* 非有限输入：本拍不判，保持锁存 / Non-finite: skip *)
        END_IF
    E_DL_HtcState.eFault:                                                      (* 故障相：冻结保持末值，仅复位沿出 / Fault *)
        ;                                                                      (* 锁存回放（R28） / Replay from latch *)
    ELSE                                                                       (* 非法相位兜底迁安全态 / Illegal phase fallback *)
        _eState := E_DL_HtcState.eFault;                                       (* 迁故障相 / To fault *)
        _bFault := TRUE;                                                       (* 同步锁存 / Latch *)
        _eCause := E_DL_HtcCause.ePhaseBad;                                    (* 成因：非法相位 / Cause: illegal phase *)
END_CASE

(* —— 段 5：出口映射（bError/eState 同源，R191） —— *)
bError := _bFault;                                                             (* 故障标志镜像 / Fault flag mirror *)
eState := _eState;                                                             (* 状态出口 / State outlet *)
eCause := _eCause;                                                             (* 成因出口 / Cause outlet *)
END_FUNCTION_BLOCK
